// LS Electric XG5000 project: SEMICON_SORTER
// PLC DR32H

PROGRAM SIM_IO (task: 스캔 프로그램)

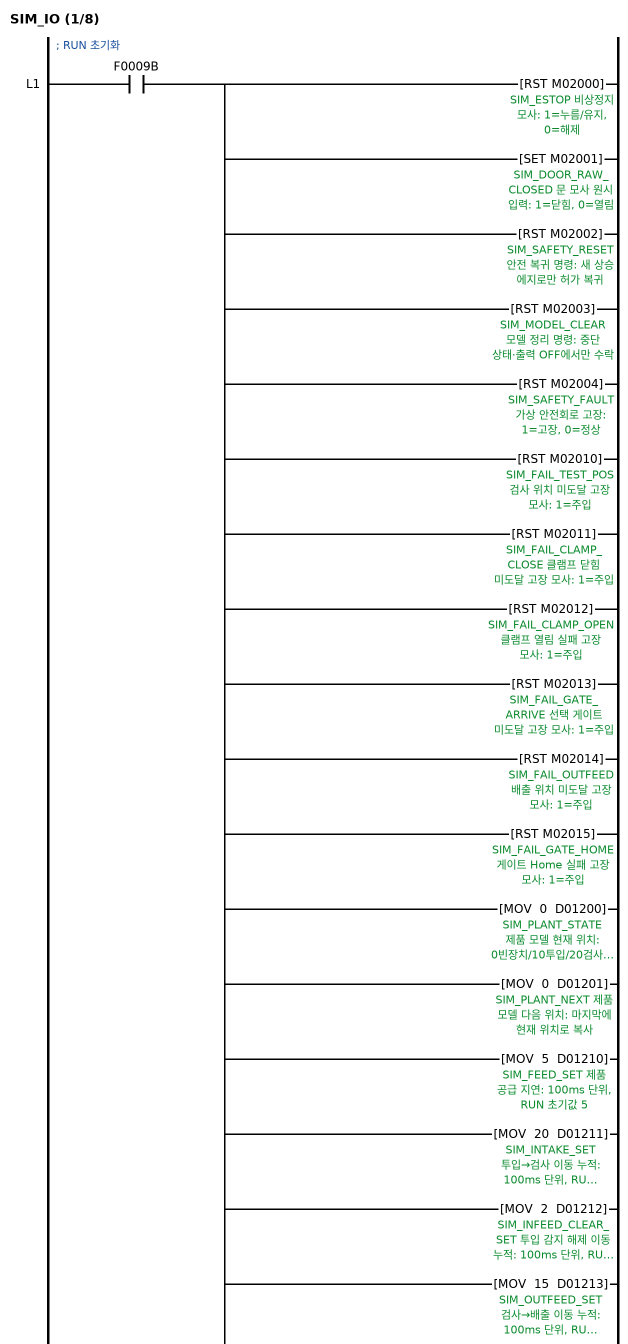

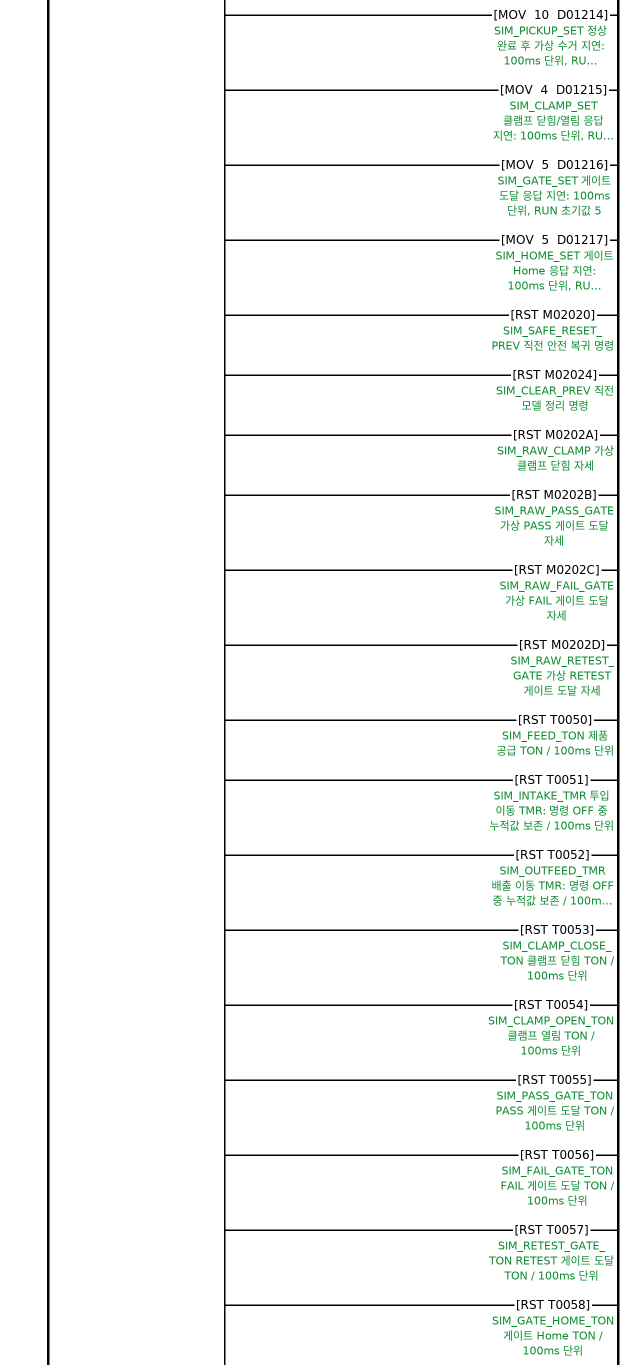

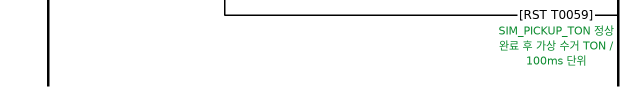
// RUN 초기화
; L1
LOAD      F0009B
RST       M02000	// SIM_ESTOP 비상정지 모사: 1=누름/유지, 0=해제
SET       M02001	// SIM_DOOR_RAW_CLOSED 문 모사 원시 입력: 1=닫힘, 0=열림
RST       M02002	// SIM_SAFETY_RESET 안전 복귀 명령: 새 상승 에지로만 허가 복귀
RST       M02003	// SIM_MODEL_CLEAR 모델 정리 명령: 중단 상태·출력 OFF에서만 수락
RST       M02004	// SIM_SAFETY_FAULT 가상 안전회로 고장: 1=고장, 0=정상
RST       M02010	// SIM_FAIL_TEST_POS 검사 위치 미도달 고장 모사: 1=주입
RST       M02011	// SIM_FAIL_CLAMP_CLOSE 클램프 닫힘 미도달 고장 모사: 1=주입
RST       M02012	// SIM_FAIL_CLAMP_OPEN 클램프 열림 실패 고장 모사: 1=주입
RST       M02013	// SIM_FAIL_GATE_ARRIVE 선택 게이트 미도달 고장 모사: 1=주입
RST       M02014	// SIM_FAIL_OUTFEED 배출 위치 미도달 고장 모사: 1=주입
RST       M02015	// SIM_FAIL_GATE_HOME 게이트 Home 실패 고장 모사: 1=주입
MOV       0 D01200	// SIM_PLANT_STATE 제품 모델 현재 위치: 0빈장치/10투입/20검사/30배출이송/40배출
MOV       0 D01201	// SIM_PLANT_NEXT 제품 모델 다음 위치: 마지막에 현재 위치로 복사
MOV       5 D01210	// SIM_FEED_SET 제품 공급 지연: 100ms 단위, RUN 초기값 5
MOV       20 D01211	// SIM_INTAKE_SET 투입→검사 이동 누적: 100ms 단위, RUN 초기값 20
MOV       2 D01212	// SIM_INFEED_CLEAR_SET 투입 감지 해제 이동 누적: 100ms 단위, RUN 초기값 2
MOV       15 D01213	// SIM_OUTFEED_SET 검사→배출 이동 누적: 100ms 단위, RUN 초기값 15
MOV       10 D01214	// SIM_PICKUP_SET 정상 완료 후 가상 수거 지연: 100ms 단위, RUN 초기값 10
MOV       4 D01215	// SIM_CLAMP_SET 클램프 닫힘/열림 응답 지연: 100ms 단위, RUN 초기값 4
MOV       5 D01216	// SIM_GATE_SET 게이트 도달 응답 지연: 100ms 단위, RUN 초기값 5
MOV       5 D01217	// SIM_HOME_SET 게이트 Home 응답 지연: 100ms 단위, RUN 초기값 5
RST       M02020	// SIM_SAFE_RESET_PREV 직전 안전 복귀 명령
RST       M02024	// SIM_CLEAR_PREV 직전 모델 정리 명령
RST       M0202A	// SIM_RAW_CLAMP 가상 클램프 닫힘 자세
RST       M0202B	// SIM_RAW_PASS_GATE 가상 PASS 게이트 도달 자세
RST       M0202C	// SIM_RAW_FAIL_GATE 가상 FAIL 게이트 도달 자세
RST       M0202D	// SIM_RAW_RETEST_GATE 가상 RETEST 게이트 도달 자세
RST       T0050	// SIM_FEED_TON 제품 공급 TON / 100ms 단위
RST       T0051	// SIM_INTAKE_TMR 투입 이동 TMR: 명령 OFF 중 누적값 보존 / 100ms 단위
RST       T0052	// SIM_OUTFEED_TMR 배출 이동 TMR: 명령 OFF 중 누적값 보존 / 100ms 단위
RST       T0053	// SIM_CLAMP_CLOSE_TON 클램프 닫힘 TON / 100ms 단위
RST       T0054	// SIM_CLAMP_OPEN_TON 클램프 열림 TON / 100ms 단위
RST       T0055	// SIM_PASS_GATE_TON PASS 게이트 도달 TON / 100ms 단위
RST       T0056	// SIM_FAIL_GATE_TON FAIL 게이트 도달 TON / 100ms 단위
RST       T0057	// SIM_RETEST_GATE_TON RETEST 게이트 도달 TON / 100ms 단위
RST       T0058	// SIM_GATE_HOME_TON 게이트 Home TON / 100ms 단위
RST       T0059	// SIM_PICKUP_TON 정상 완료 후 가상 수거 TON / 100ms 단위

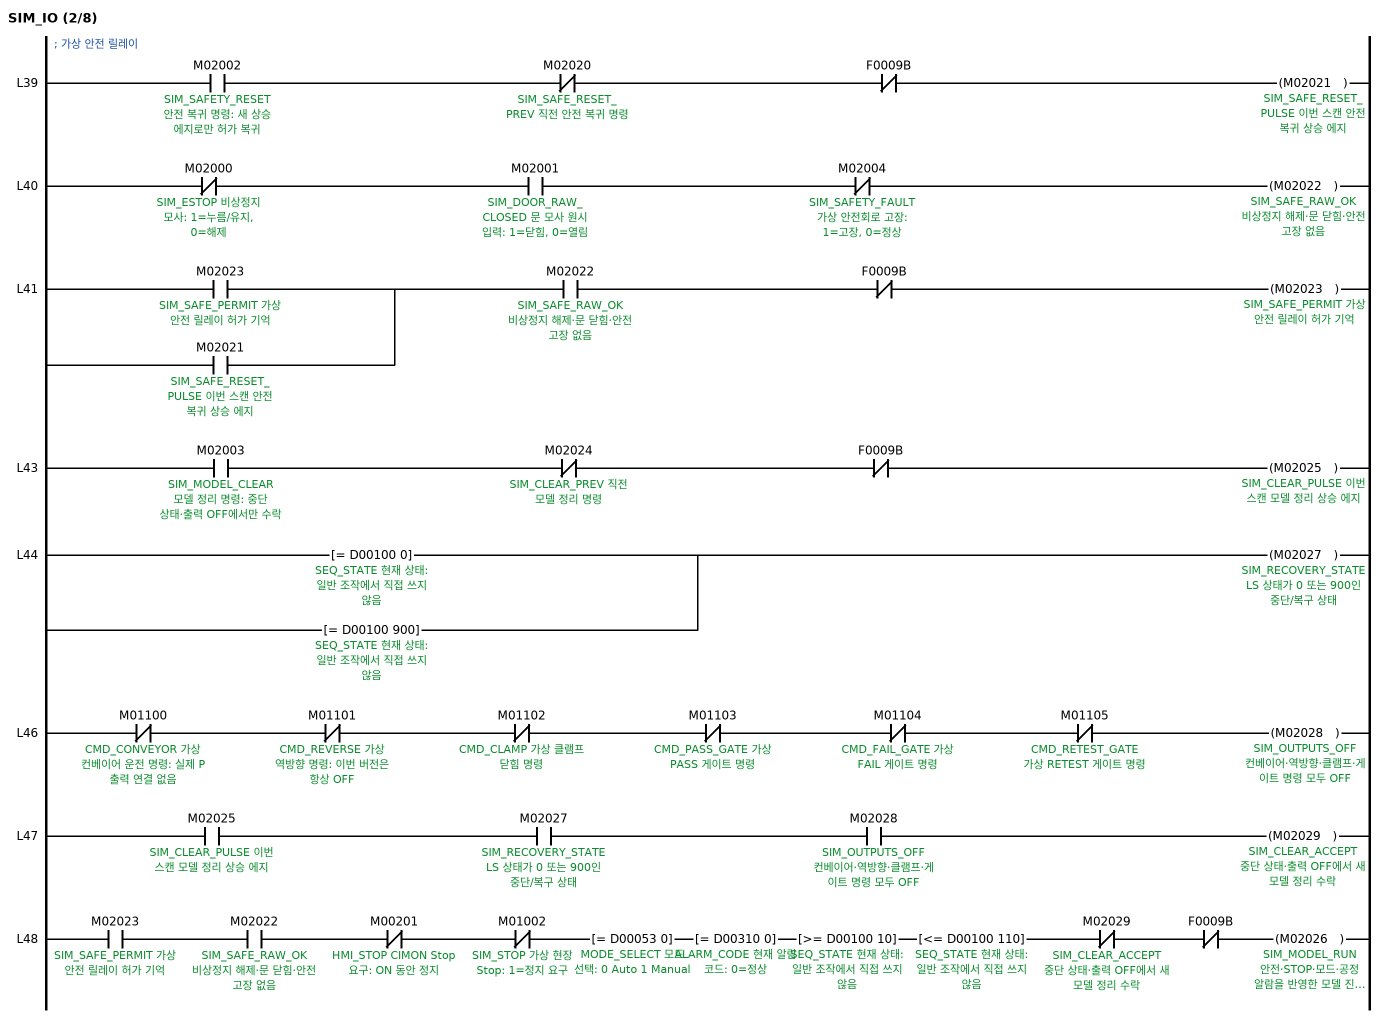
// 가상 안전 릴레이
; L39
LOAD      M02002	// SIM_SAFETY_RESET 안전 복귀 명령: 새 상승 에지로만 허가 복귀
AND NOT   M02020	// SIM_SAFE_RESET_PREV 직전 안전 복귀 명령
AND NOT   F0009B
OUT       M02021	// SIM_SAFE_RESET_PULSE 이번 스캔 안전 복귀 상승 에지
; L40
LOAD NOT  M02000	// SIM_ESTOP 비상정지 모사: 1=누름/유지, 0=해제
AND       M02001	// SIM_DOOR_RAW_CLOSED 문 모사 원시 입력: 1=닫힘, 0=열림
AND NOT   M02004	// SIM_SAFETY_FAULT 가상 안전회로 고장: 1=고장, 0=정상
OUT       M02022	// SIM_SAFE_RAW_OK 비상정지 해제·문 닫힘·안전 고장 없음
; L41
LOAD      M02023	// SIM_SAFE_PERMIT 가상 안전 릴레이 허가 기억
OR        M02021	// SIM_SAFE_RESET_PULSE 이번 스캔 안전 복귀 상승 에지
AND       M02022	// SIM_SAFE_RAW_OK 비상정지 해제·문 닫힘·안전 고장 없음
AND NOT   F0009B
OUT       M02023	// SIM_SAFE_PERMIT 가상 안전 릴레이 허가 기억
; L43
LOAD      M02003	// SIM_MODEL_CLEAR 모델 정리 명령: 중단 상태·출력 OFF에서만 수락
AND NOT   M02024	// SIM_CLEAR_PREV 직전 모델 정리 명령
AND NOT   F0009B
OUT       M02025	// SIM_CLEAR_PULSE 이번 스캔 모델 정리 상승 에지
; L44
LOAD=     D00100 0	// SEQ_STATE 현재 상태: 일반 조작에서 직접 쓰지 않음
OR=       D00100 900	// SEQ_STATE 현재 상태: 일반 조작에서 직접 쓰지 않음
OUT       M02027	// SIM_RECOVERY_STATE LS 상태가 0 또는 900인 중단/복구 상태
; L46
LOAD NOT  M01100	// CMD_CONVEYOR 가상 컨베이어 운전 명령: 실제 P 출력 연결 없음
AND NOT   M01101	// CMD_REVERSE 가상 역방향 명령: 이번 버전은 항상 OFF
AND NOT   M01102	// CMD_CLAMP 가상 클램프 닫힘 명령
AND NOT   M01103	// CMD_PASS_GATE 가상 PASS 게이트 명령
AND NOT   M01104	// CMD_FAIL_GATE 가상 FAIL 게이트 명령
AND NOT   M01105	// CMD_RETEST_GATE 가상 RETEST 게이트 명령
OUT       M02028	// SIM_OUTPUTS_OFF 컨베이어·역방향·클램프·게이트 명령 모두 OFF
; L47
LOAD      M02025	// SIM_CLEAR_PULSE 이번 스캔 모델 정리 상승 에지
AND       M02027	// SIM_RECOVERY_STATE LS 상태가 0 또는 900인 중단/복구 상태
AND       M02028	// SIM_OUTPUTS_OFF 컨베이어·역방향·클램프·게이트 명령 모두 OFF
OUT       M02029	// SIM_CLEAR_ACCEPT 중단 상태·출력 OFF에서 새 모델 정리 수락
; L48
LOAD      M02023	// SIM_SAFE_PERMIT 가상 안전 릴레이 허가 기억
AND       M02022	// SIM_SAFE_RAW_OK 비상정지 해제·문 닫힘·안전 고장 없음
AND NOT   M00201	// HMI_STOP CIMON Stop 요구: ON 동안 정지
AND NOT   M01002	// SIM_STOP 가상 현장 Stop: 1=정지 요구
AND=      D00053 0	// MODE_SELECT 모드 선택: 0 Auto 1 Manual
AND=      D00310 0	// ALARM_CODE 현재 알람 코드: 0=정상
AND>=     D00100 10	// SEQ_STATE 현재 상태: 일반 조작에서 직접 쓰지 않음
AND<=     D00100 110	// SEQ_STATE 현재 상태: 일반 조작에서 직접 쓰지 않음
AND NOT   M02029	// SIM_CLEAR_ACCEPT 중단 상태·출력 OFF에서 새 모델 정리 수락
AND NOT   F0009B
OUT       M02026	// SIM_MODEL_RUN 안전·STOP·모드·공정 알람을 반영한 모델 진행 허가

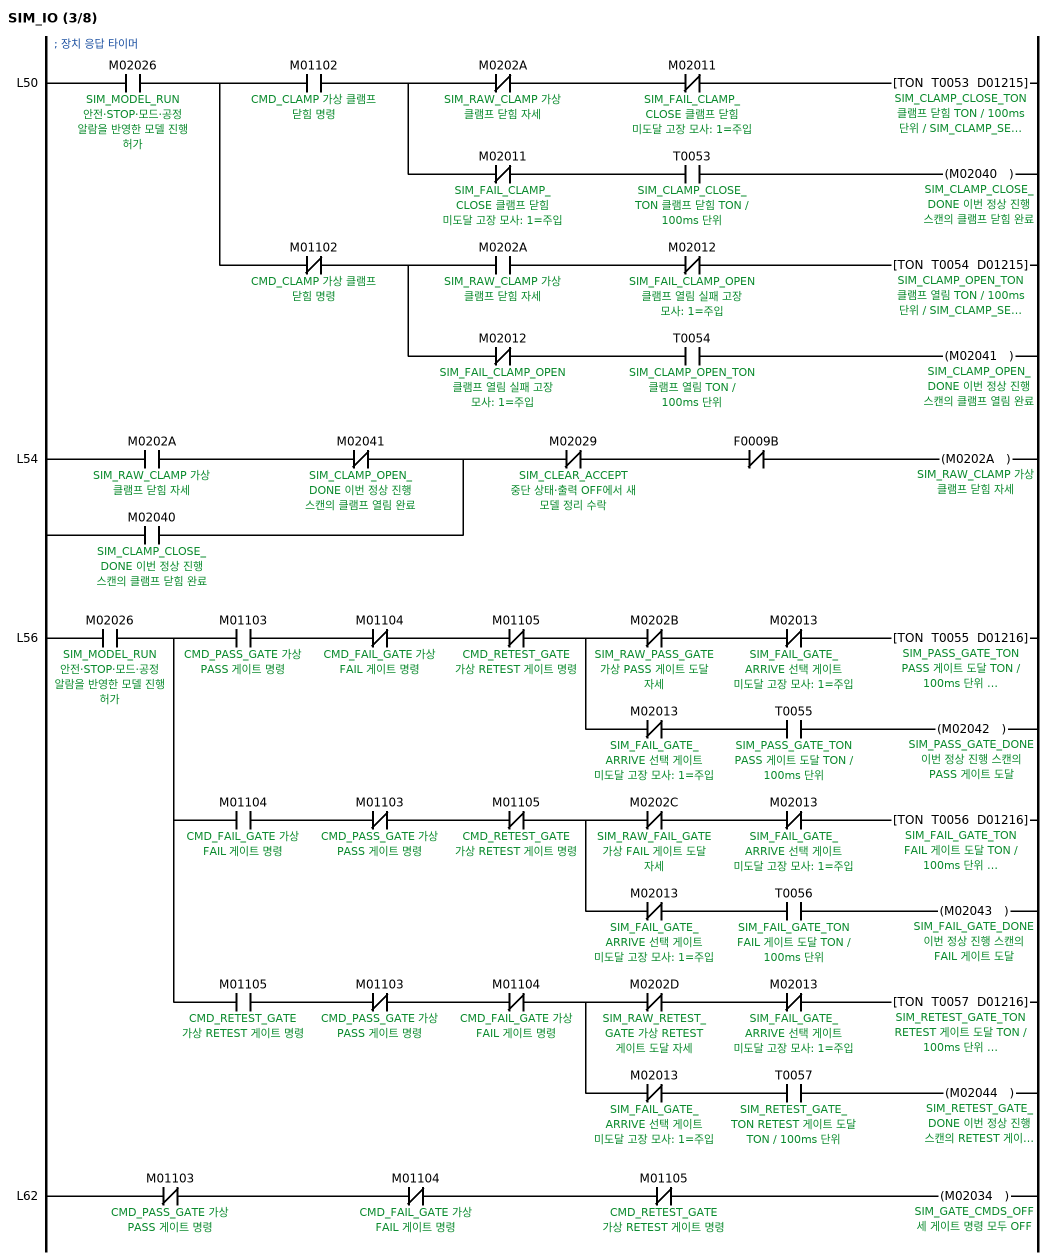
// 장치 응답 타이머
; L50
LOAD      M02026	// SIM_MODEL_RUN 안전·STOP·모드·공정 알람을 반영한 모델 진행 허가
MPUSH
AND       M01102	// CMD_CLAMP 가상 클램프 닫힘 명령
MPUSH
AND NOT   M0202A	// SIM_RAW_CLAMP 가상 클램프 닫힘 자세
AND NOT   M02011	// SIM_FAIL_CLAMP_CLOSE 클램프 닫힘 미도달 고장 모사: 1=주입
TON       T0053 D01215	// SIM_CLAMP_CLOSE_TON 클램프 닫힘 TON / 100ms 단위 / SIM_CLAMP_SET 클램프 닫힘/열림 응답 지연: 100ms 단위, RUN 초기값 4
MPOP
AND NOT   M02011	// SIM_FAIL_CLAMP_CLOSE 클램프 닫힘 미도달 고장 모사: 1=주입
AND       T0053	// SIM_CLAMP_CLOSE_TON 클램프 닫힘 TON / 100ms 단위
OUT       M02040	// SIM_CLAMP_CLOSE_DONE 이번 정상 진행 스캔의 클램프 닫힘 완료
MPOP
AND NOT   M01102	// CMD_CLAMP 가상 클램프 닫힘 명령
MPUSH
AND       M0202A	// SIM_RAW_CLAMP 가상 클램프 닫힘 자세
AND NOT   M02012	// SIM_FAIL_CLAMP_OPEN 클램프 열림 실패 고장 모사: 1=주입
TON       T0054 D01215	// SIM_CLAMP_OPEN_TON 클램프 열림 TON / 100ms 단위 / SIM_CLAMP_SET 클램프 닫힘/열림 응답 지연: 100ms 단위, RUN 초기값 4
MPOP
AND NOT   M02012	// SIM_FAIL_CLAMP_OPEN 클램프 열림 실패 고장 모사: 1=주입
AND       T0054	// SIM_CLAMP_OPEN_TON 클램프 열림 TON / 100ms 단위
OUT       M02041	// SIM_CLAMP_OPEN_DONE 이번 정상 진행 스캔의 클램프 열림 완료
; L54
LOAD      M0202A	// SIM_RAW_CLAMP 가상 클램프 닫힘 자세
AND NOT   M02041	// SIM_CLAMP_OPEN_DONE 이번 정상 진행 스캔의 클램프 열림 완료
OR        M02040	// SIM_CLAMP_CLOSE_DONE 이번 정상 진행 스캔의 클램프 닫힘 완료
AND NOT   M02029	// SIM_CLEAR_ACCEPT 중단 상태·출력 OFF에서 새 모델 정리 수락
AND NOT   F0009B
OUT       M0202A	// SIM_RAW_CLAMP 가상 클램프 닫힘 자세
; L56
LOAD      M02026	// SIM_MODEL_RUN 안전·STOP·모드·공정 알람을 반영한 모델 진행 허가
MPUSH
AND       M01103	// CMD_PASS_GATE 가상 PASS 게이트 명령
AND NOT   M01104	// CMD_FAIL_GATE 가상 FAIL 게이트 명령
AND NOT   M01105	// CMD_RETEST_GATE 가상 RETEST 게이트 명령
MPUSH
AND NOT   M0202B	// SIM_RAW_PASS_GATE 가상 PASS 게이트 도달 자세
AND NOT   M02013	// SIM_FAIL_GATE_ARRIVE 선택 게이트 미도달 고장 모사: 1=주입
TON       T0055 D01216	// SIM_PASS_GATE_TON PASS 게이트 도달 TON / 100ms 단위 / SIM_GATE_SET 게이트 도달 응답 지연: 100ms 단위, RUN 초기값 5
MPOP
AND NOT   M02013	// SIM_FAIL_GATE_ARRIVE 선택 게이트 미도달 고장 모사: 1=주입
AND       T0055	// SIM_PASS_GATE_TON PASS 게이트 도달 TON / 100ms 단위
OUT       M02042	// SIM_PASS_GATE_DONE 이번 정상 진행 스캔의 PASS 게이트 도달
MLOAD
AND       M01104	// CMD_FAIL_GATE 가상 FAIL 게이트 명령
AND NOT   M01103	// CMD_PASS_GATE 가상 PASS 게이트 명령
AND NOT   M01105	// CMD_RETEST_GATE 가상 RETEST 게이트 명령
MPUSH
AND NOT   M0202C	// SIM_RAW_FAIL_GATE 가상 FAIL 게이트 도달 자세
AND NOT   M02013	// SIM_FAIL_GATE_ARRIVE 선택 게이트 미도달 고장 모사: 1=주입
TON       T0056 D01216	// SIM_FAIL_GATE_TON FAIL 게이트 도달 TON / 100ms 단위 / SIM_GATE_SET 게이트 도달 응답 지연: 100ms 단위, RUN 초기값 5
MPOP
AND NOT   M02013	// SIM_FAIL_GATE_ARRIVE 선택 게이트 미도달 고장 모사: 1=주입
AND       T0056	// SIM_FAIL_GATE_TON FAIL 게이트 도달 TON / 100ms 단위
OUT       M02043	// SIM_FAIL_GATE_DONE 이번 정상 진행 스캔의 FAIL 게이트 도달
MPOP
AND       M01105	// CMD_RETEST_GATE 가상 RETEST 게이트 명령
AND NOT   M01103	// CMD_PASS_GATE 가상 PASS 게이트 명령
AND NOT   M01104	// CMD_FAIL_GATE 가상 FAIL 게이트 명령
MPUSH
AND NOT   M0202D	// SIM_RAW_RETEST_GATE 가상 RETEST 게이트 도달 자세
AND NOT   M02013	// SIM_FAIL_GATE_ARRIVE 선택 게이트 미도달 고장 모사: 1=주입
TON       T0057 D01216	// SIM_RETEST_GATE_TON RETEST 게이트 도달 TON / 100ms 단위 / SIM_GATE_SET 게이트 도달 응답 지연: 100ms 단위, RUN 초기값 5
MPOP
AND NOT   M02013	// SIM_FAIL_GATE_ARRIVE 선택 게이트 미도달 고장 모사: 1=주입
AND       T0057	// SIM_RETEST_GATE_TON RETEST 게이트 도달 TON / 100ms 단위
OUT       M02044	// SIM_RETEST_GATE_DONE 이번 정상 진행 스캔의 RETEST 게이트 도달
; L62
LOAD NOT  M01103	// CMD_PASS_GATE 가상 PASS 게이트 명령
AND NOT   M01104	// CMD_FAIL_GATE 가상 FAIL 게이트 명령
AND NOT   M01105	// CMD_RETEST_GATE 가상 RETEST 게이트 명령
OUT       M02034	// SIM_GATE_CMDS_OFF 세 게이트 명령 모두 OFF

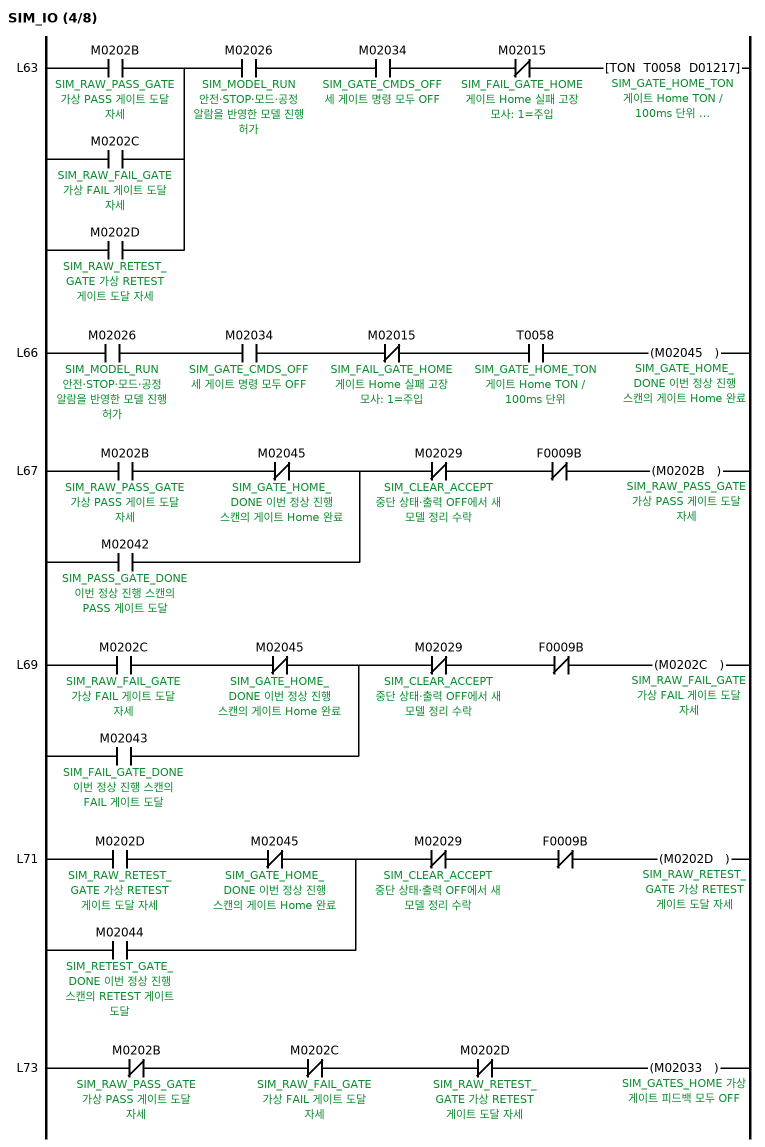
; L63
LOAD      M0202B	// SIM_RAW_PASS_GATE 가상 PASS 게이트 도달 자세
OR        M0202C	// SIM_RAW_FAIL_GATE 가상 FAIL 게이트 도달 자세
OR        M0202D	// SIM_RAW_RETEST_GATE 가상 RETEST 게이트 도달 자세
AND       M02026	// SIM_MODEL_RUN 안전·STOP·모드·공정 알람을 반영한 모델 진행 허가
AND       M02034	// SIM_GATE_CMDS_OFF 세 게이트 명령 모두 OFF
AND NOT   M02015	// SIM_FAIL_GATE_HOME 게이트 Home 실패 고장 모사: 1=주입
TON       T0058 D01217	// SIM_GATE_HOME_TON 게이트 Home TON / 100ms 단위 / SIM_HOME_SET 게이트 Home 응답 지연: 100ms 단위, RUN 초기값 5
; L66
LOAD      M02026	// SIM_MODEL_RUN 안전·STOP·모드·공정 알람을 반영한 모델 진행 허가
AND       M02034	// SIM_GATE_CMDS_OFF 세 게이트 명령 모두 OFF
AND NOT   M02015	// SIM_FAIL_GATE_HOME 게이트 Home 실패 고장 모사: 1=주입
AND       T0058	// SIM_GATE_HOME_TON 게이트 Home TON / 100ms 단위
OUT       M02045	// SIM_GATE_HOME_DONE 이번 정상 진행 스캔의 게이트 Home 완료
; L67
LOAD      M0202B	// SIM_RAW_PASS_GATE 가상 PASS 게이트 도달 자세
AND NOT   M02045	// SIM_GATE_HOME_DONE 이번 정상 진행 스캔의 게이트 Home 완료
OR        M02042	// SIM_PASS_GATE_DONE 이번 정상 진행 스캔의 PASS 게이트 도달
AND NOT   M02029	// SIM_CLEAR_ACCEPT 중단 상태·출력 OFF에서 새 모델 정리 수락
AND NOT   F0009B
OUT       M0202B	// SIM_RAW_PASS_GATE 가상 PASS 게이트 도달 자세
; L69
LOAD      M0202C	// SIM_RAW_FAIL_GATE 가상 FAIL 게이트 도달 자세
AND NOT   M02045	// SIM_GATE_HOME_DONE 이번 정상 진행 스캔의 게이트 Home 완료
OR        M02043	// SIM_FAIL_GATE_DONE 이번 정상 진행 스캔의 FAIL 게이트 도달
AND NOT   M02029	// SIM_CLEAR_ACCEPT 중단 상태·출력 OFF에서 새 모델 정리 수락
AND NOT   F0009B
OUT       M0202C	// SIM_RAW_FAIL_GATE 가상 FAIL 게이트 도달 자세
; L71
LOAD      M0202D	// SIM_RAW_RETEST_GATE 가상 RETEST 게이트 도달 자세
AND NOT   M02045	// SIM_GATE_HOME_DONE 이번 정상 진행 스캔의 게이트 Home 완료
OR        M02044	// SIM_RETEST_GATE_DONE 이번 정상 진행 스캔의 RETEST 게이트 도달
AND NOT   M02029	// SIM_CLEAR_ACCEPT 중단 상태·출력 OFF에서 새 모델 정리 수락
AND NOT   F0009B
OUT       M0202D	// SIM_RAW_RETEST_GATE 가상 RETEST 게이트 도달 자세
; L73
LOAD NOT  M0202B	// SIM_RAW_PASS_GATE 가상 PASS 게이트 도달 자세
AND NOT   M0202C	// SIM_RAW_FAIL_GATE 가상 FAIL 게이트 도달 자세
AND NOT   M0202D	// SIM_RAW_RETEST_GATE 가상 RETEST 게이트 도달 자세
OUT       M02033	// SIM_GATES_HOME 가상 게이트 피드백 모두 OFF

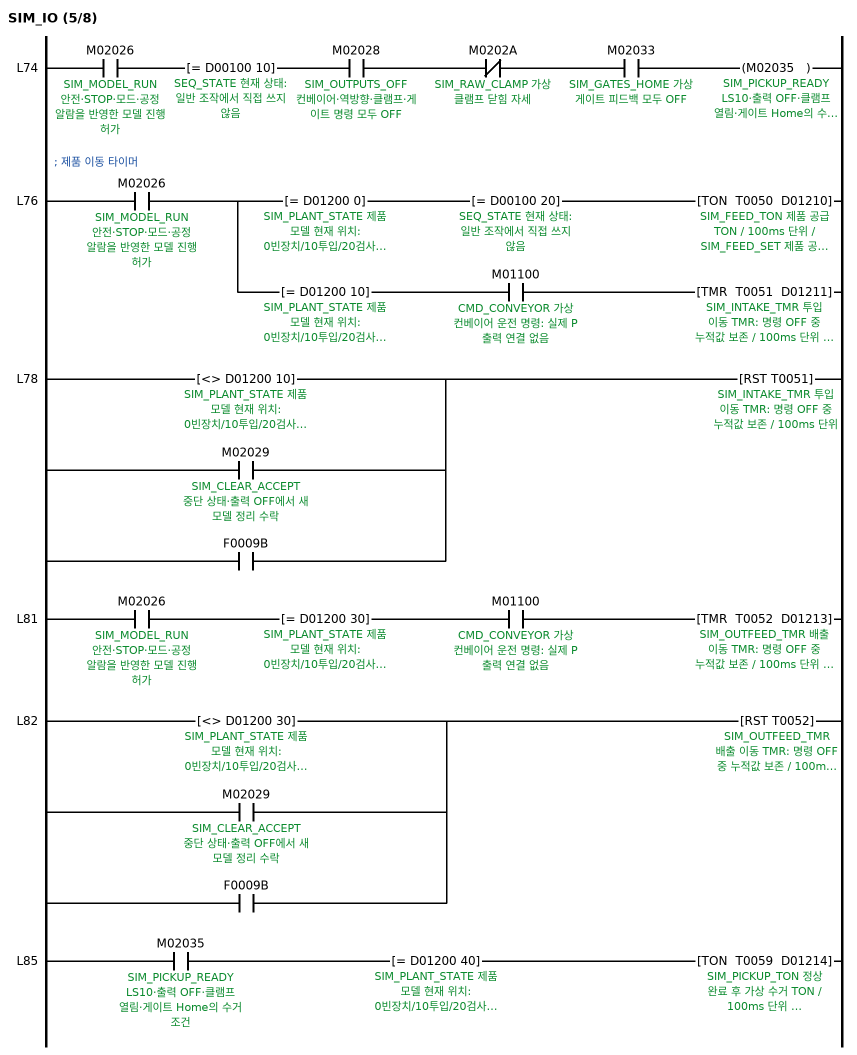
; L74
LOAD      M02026	// SIM_MODEL_RUN 안전·STOP·모드·공정 알람을 반영한 모델 진행 허가
AND=      D00100 10	// SEQ_STATE 현재 상태: 일반 조작에서 직접 쓰지 않음
AND       M02028	// SIM_OUTPUTS_OFF 컨베이어·역방향·클램프·게이트 명령 모두 OFF
AND NOT   M0202A	// SIM_RAW_CLAMP 가상 클램프 닫힘 자세
AND       M02033	// SIM_GATES_HOME 가상 게이트 피드백 모두 OFF
OUT       M02035	// SIM_PICKUP_READY LS10·출력 OFF·클램프 열림·게이트 Home의 수거 조건
// 제품 이동 타이머
; L76
LOAD      M02026	// SIM_MODEL_RUN 안전·STOP·모드·공정 알람을 반영한 모델 진행 허가
MPUSH
AND=      D01200 0	// SIM_PLANT_STATE 제품 모델 현재 위치: 0빈장치/10투입/20검사/30배출이송/40배출
AND=      D00100 20	// SEQ_STATE 현재 상태: 일반 조작에서 직접 쓰지 않음
TON       T0050 D01210	// SIM_FEED_TON 제품 공급 TON / 100ms 단위 / SIM_FEED_SET 제품 공급 지연: 100ms 단위, RUN 초기값 5
MPOP
AND=      D01200 10	// SIM_PLANT_STATE 제품 모델 현재 위치: 0빈장치/10투입/20검사/30배출이송/40배출
AND       M01100	// CMD_CONVEYOR 가상 컨베이어 운전 명령: 실제 P 출력 연결 없음
TMR       T0051 D01211	// SIM_INTAKE_TMR 투입 이동 TMR: 명령 OFF 중 누적값 보존 / 100ms 단위 / SIM_INTAKE_SET 투입→검사 이동 누적: 100ms 단위, RUN 초기값 20
; L78
LOAD<>    D01200 10	// SIM_PLANT_STATE 제품 모델 현재 위치: 0빈장치/10투입/20검사/30배출이송/40배출
OR        M02029	// SIM_CLEAR_ACCEPT 중단 상태·출력 OFF에서 새 모델 정리 수락
OR        F0009B
RST       T0051	// SIM_INTAKE_TMR 투입 이동 TMR: 명령 OFF 중 누적값 보존 / 100ms 단위
; L81
LOAD      M02026	// SIM_MODEL_RUN 안전·STOP·모드·공정 알람을 반영한 모델 진행 허가
AND=      D01200 30	// SIM_PLANT_STATE 제품 모델 현재 위치: 0빈장치/10투입/20검사/30배출이송/40배출
AND       M01100	// CMD_CONVEYOR 가상 컨베이어 운전 명령: 실제 P 출력 연결 없음
TMR       T0052 D01213	// SIM_OUTFEED_TMR 배출 이동 TMR: 명령 OFF 중 누적값 보존 / 100ms 단위 / SIM_OUTFEED_SET 검사→배출 이동 누적: 100ms 단위, RUN 초기값 15
; L82
LOAD<>    D01200 30	// SIM_PLANT_STATE 제품 모델 현재 위치: 0빈장치/10투입/20검사/30배출이송/40배출
OR        M02029	// SIM_CLEAR_ACCEPT 중단 상태·출력 OFF에서 새 모델 정리 수락
OR        F0009B
RST       T0052	// SIM_OUTFEED_TMR 배출 이동 TMR: 명령 OFF 중 누적값 보존 / 100ms 단위
; L85
LOAD      M02035	// SIM_PICKUP_READY LS10·출력 OFF·클램프 열림·게이트 Home의 수거 조건
AND=      D01200 40	// SIM_PLANT_STATE 제품 모델 현재 위치: 0빈장치/10투입/20검사/30배출이송/40배출
TON       T0059 D01214	// SIM_PICKUP_TON 정상 완료 후 가상 수거 TON / 100ms 단위 / SIM_PICKUP_SET 정상 완료 후 가상 수거 지연: 100ms 단위, RUN 초기값 10

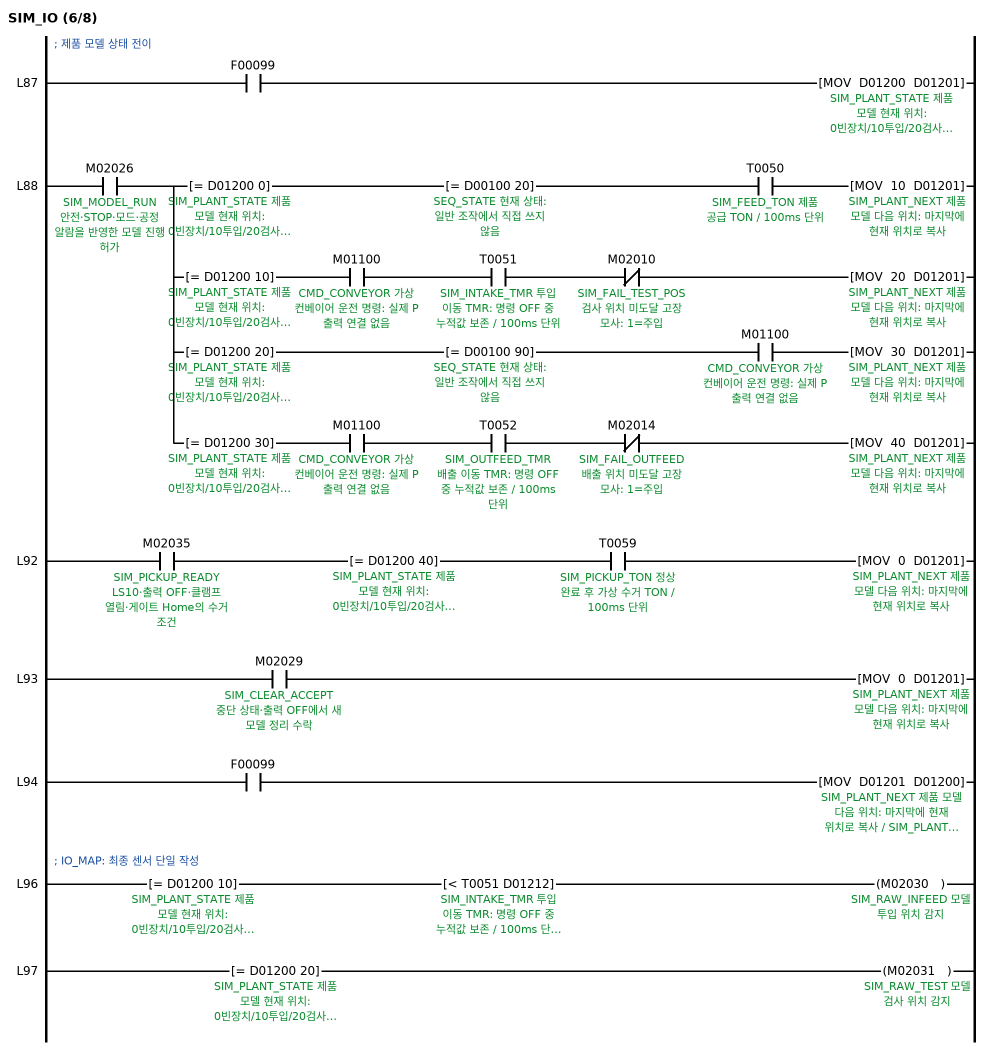
// 제품 모델 상태 전이
; L87
LOAD      F00099
MOV       D01200 D01201	// SIM_PLANT_STATE 제품 모델 현재 위치: 0빈장치/10투입/20검사/30배출이송/40배출 / SIM_PLANT_NEXT 제품 모델 다음 위치: 마지막에 현재 위치로 복사
; L88
LOAD      M02026	// SIM_MODEL_RUN 안전·STOP·모드·공정 알람을 반영한 모델 진행 허가
MPUSH
AND=      D01200 0	// SIM_PLANT_STATE 제품 모델 현재 위치: 0빈장치/10투입/20검사/30배출이송/40배출
AND=      D00100 20	// SEQ_STATE 현재 상태: 일반 조작에서 직접 쓰지 않음
AND       T0050	// SIM_FEED_TON 제품 공급 TON / 100ms 단위
MOV       10 D01201	// SIM_PLANT_NEXT 제품 모델 다음 위치: 마지막에 현재 위치로 복사
MLOAD
AND=      D01200 10	// SIM_PLANT_STATE 제품 모델 현재 위치: 0빈장치/10투입/20검사/30배출이송/40배출
AND       M01100	// CMD_CONVEYOR 가상 컨베이어 운전 명령: 실제 P 출력 연결 없음
AND       T0051	// SIM_INTAKE_TMR 투입 이동 TMR: 명령 OFF 중 누적값 보존 / 100ms 단위
AND NOT   M02010	// SIM_FAIL_TEST_POS 검사 위치 미도달 고장 모사: 1=주입
MOV       20 D01201	// SIM_PLANT_NEXT 제품 모델 다음 위치: 마지막에 현재 위치로 복사
MLOAD
AND=      D01200 20	// SIM_PLANT_STATE 제품 모델 현재 위치: 0빈장치/10투입/20검사/30배출이송/40배출
AND=      D00100 90	// SEQ_STATE 현재 상태: 일반 조작에서 직접 쓰지 않음
AND       M01100	// CMD_CONVEYOR 가상 컨베이어 운전 명령: 실제 P 출력 연결 없음
MOV       30 D01201	// SIM_PLANT_NEXT 제품 모델 다음 위치: 마지막에 현재 위치로 복사
MPOP
AND=      D01200 30	// SIM_PLANT_STATE 제품 모델 현재 위치: 0빈장치/10투입/20검사/30배출이송/40배출
AND       M01100	// CMD_CONVEYOR 가상 컨베이어 운전 명령: 실제 P 출력 연결 없음
AND       T0052	// SIM_OUTFEED_TMR 배출 이동 TMR: 명령 OFF 중 누적값 보존 / 100ms 단위
AND NOT   M02014	// SIM_FAIL_OUTFEED 배출 위치 미도달 고장 모사: 1=주입
MOV       40 D01201	// SIM_PLANT_NEXT 제품 모델 다음 위치: 마지막에 현재 위치로 복사
; L92
LOAD      M02035	// SIM_PICKUP_READY LS10·출력 OFF·클램프 열림·게이트 Home의 수거 조건
AND=      D01200 40	// SIM_PLANT_STATE 제품 모델 현재 위치: 0빈장치/10투입/20검사/30배출이송/40배출
AND       T0059	// SIM_PICKUP_TON 정상 완료 후 가상 수거 TON / 100ms 단위
MOV       0 D01201	// SIM_PLANT_NEXT 제품 모델 다음 위치: 마지막에 현재 위치로 복사
; L93
LOAD      M02029	// SIM_CLEAR_ACCEPT 중단 상태·출력 OFF에서 새 모델 정리 수락
MOV       0 D01201	// SIM_PLANT_NEXT 제품 모델 다음 위치: 마지막에 현재 위치로 복사
; L94
LOAD      F00099
MOV       D01201 D01200	// SIM_PLANT_NEXT 제품 모델 다음 위치: 마지막에 현재 위치로 복사 / SIM_PLANT_STATE 제품 모델 현재 위치: 0빈장치/10투입/20검사/30배출이송/40배출
// IO_MAP: 최종 센서 단일 작성
; L96
LOAD=     D01200 10	// SIM_PLANT_STATE 제품 모델 현재 위치: 0빈장치/10투입/20검사/30배출이송/40배출
AND<      T0051 D01212	// SIM_INTAKE_TMR 투입 이동 TMR: 명령 OFF 중 누적값 보존 / 100ms 단위 / SIM_INFEED_CLEAR_SET 투입 감지 해제 이동 누적: 100ms 단위, RUN 초기값 2
OUT       M02030	// SIM_RAW_INFEED 모델 투입 위치 감지
; L97
LOAD=     D01200 20	// SIM_PLANT_STATE 제품 모델 현재 위치: 0빈장치/10투입/20검사/30배출이송/40배출
OUT       M02031	// SIM_RAW_TEST 모델 검사 위치 감지

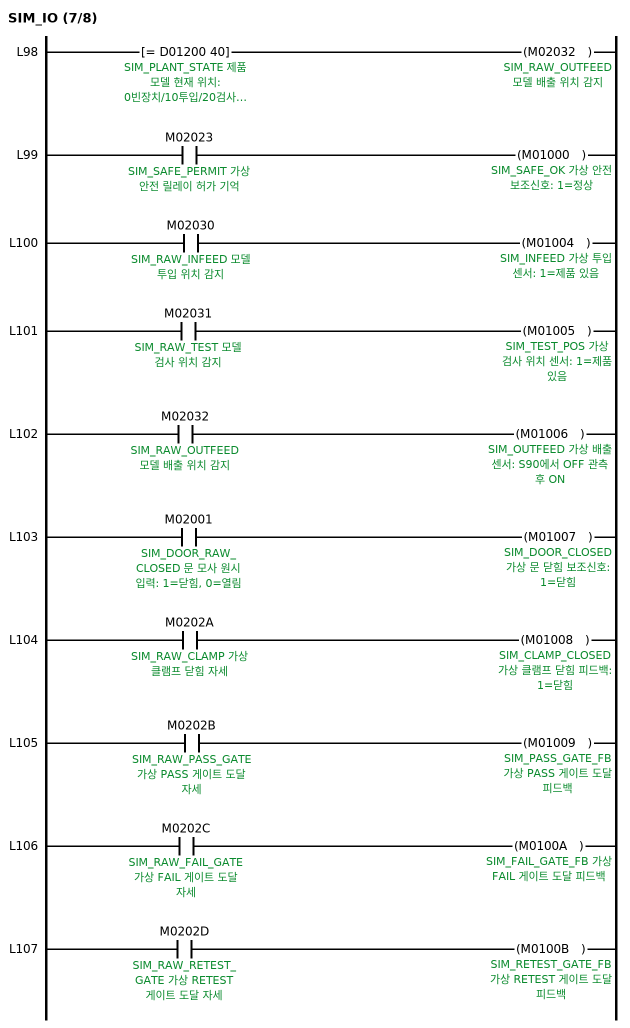
; L98
LOAD=     D01200 40	// SIM_PLANT_STATE 제품 모델 현재 위치: 0빈장치/10투입/20검사/30배출이송/40배출
OUT       M02032	// SIM_RAW_OUTFEED 모델 배출 위치 감지
; L99
LOAD      M02023	// SIM_SAFE_PERMIT 가상 안전 릴레이 허가 기억
OUT       M01000	// SIM_SAFE_OK 가상 안전 보조신호: 1=정상
; L100
LOAD      M02030	// SIM_RAW_INFEED 모델 투입 위치 감지
OUT       M01004	// SIM_INFEED 가상 투입 센서: 1=제품 있음
; L101
LOAD      M02031	// SIM_RAW_TEST 모델 검사 위치 감지
OUT       M01005	// SIM_TEST_POS 가상 검사 위치 센서: 1=제품 있음
; L102
LOAD      M02032	// SIM_RAW_OUTFEED 모델 배출 위치 감지
OUT       M01006	// SIM_OUTFEED 가상 배출 센서: S90에서 OFF 관측 후 ON
; L103
LOAD      M02001	// SIM_DOOR_RAW_CLOSED 문 모사 원시 입력: 1=닫힘, 0=열림
OUT       M01007	// SIM_DOOR_CLOSED 가상 문 닫힘 보조신호: 1=닫힘
; L104
LOAD      M0202A	// SIM_RAW_CLAMP 가상 클램프 닫힘 자세
OUT       M01008	// SIM_CLAMP_CLOSED 가상 클램프 닫힘 피드백: 1=닫힘
; L105
LOAD      M0202B	// SIM_RAW_PASS_GATE 가상 PASS 게이트 도달 자세
OUT       M01009	// SIM_PASS_GATE_FB 가상 PASS 게이트 도달 피드백
; L106
LOAD      M0202C	// SIM_RAW_FAIL_GATE 가상 FAIL 게이트 도달 자세
OUT       M0100A	// SIM_FAIL_GATE_FB 가상 FAIL 게이트 도달 피드백
; L107
LOAD      M0202D	// SIM_RAW_RETEST_GATE 가상 RETEST 게이트 도달 자세
OUT       M0100B	// SIM_RETEST_GATE_FB 가상 RETEST 게이트 도달 피드백

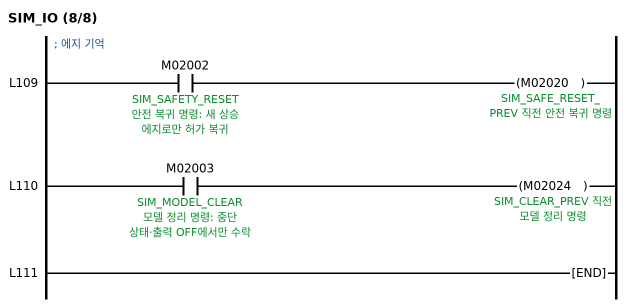
// 에지 기억
; L109
LOAD      M02002	// SIM_SAFETY_RESET 안전 복귀 명령: 새 상승 에지로만 허가 복귀
OUT       M02020	// SIM_SAFE_RESET_PREV 직전 안전 복귀 명령
; L110
LOAD      M02003	// SIM_MODEL_CLEAR 모델 정리 명령: 중단 상태·출력 OFF에서만 수락
OUT       M02024	// SIM_CLEAR_PREV 직전 모델 정리 명령
; L111
END

PROGRAM MAIN (task: 스캔 프로그램)

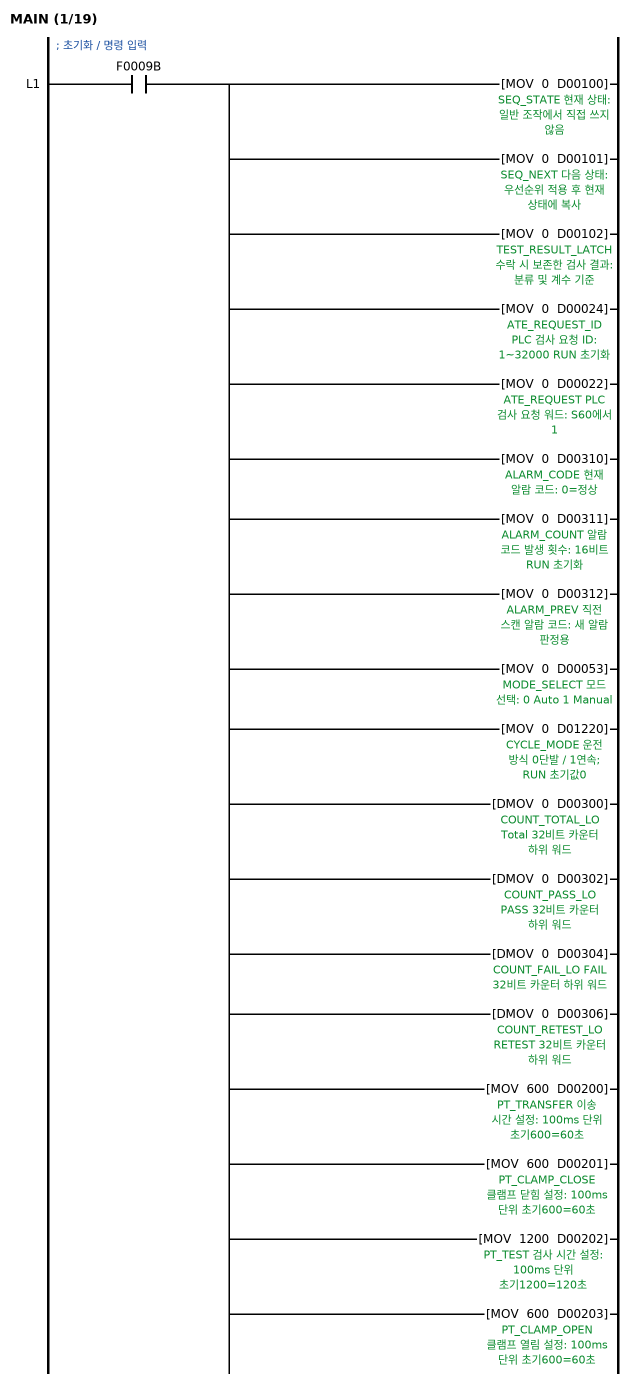

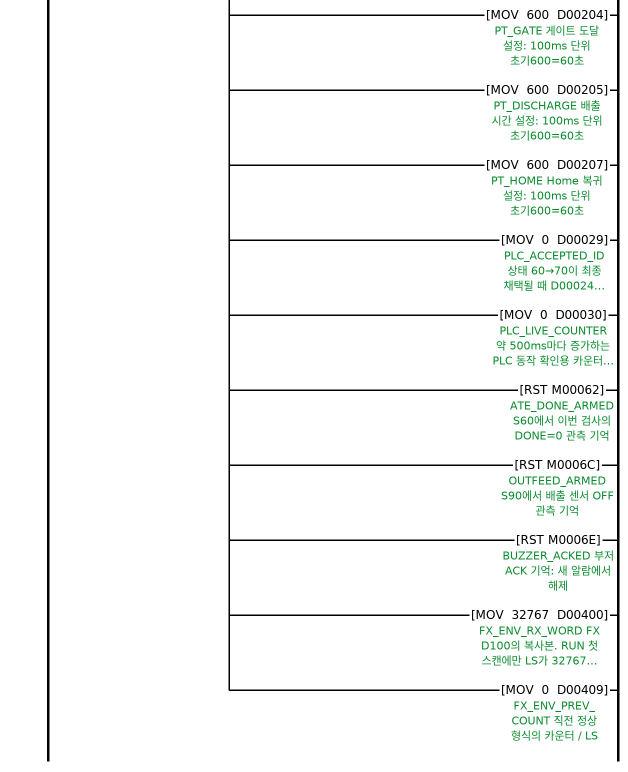
// 초기화 / 명령 입력
; L1
LOAD      F0009B
MOV       0 D00100	// SEQ_STATE 현재 상태: 일반 조작에서 직접 쓰지 않음
MOV       0 D00101	// SEQ_NEXT 다음 상태: 우선순위 적용 후 현재 상태에 복사
MOV       0 D00102	// TEST_RESULT_LATCH 수락 시 보존한 검사 결과: 분류 및 계수 기준
MOV       0 D00024	// ATE_REQUEST_ID PLC 검사 요청 ID: 1~32000 RUN 초기화
MOV       0 D00022	// ATE_REQUEST PLC 검사 요청 워드: S60에서 1
MOV       0 D00310	// ALARM_CODE 현재 알람 코드: 0=정상
MOV       0 D00311	// ALARM_COUNT 알람 코드 발생 횟수: 16비트 RUN 초기화
MOV       0 D00312	// ALARM_PREV 직전 스캔 알람 코드: 새 알람 판정용
MOV       0 D00053	// MODE_SELECT 모드 선택: 0 Auto 1 Manual
MOV       0 D01220	// CYCLE_MODE 운전 방식 0단발 / 1연속; RUN 초기값0
DMOV      0 D00300	// COUNT_TOTAL_LO Total 32비트 카운터 하위 워드
DMOV      0 D00302	// COUNT_PASS_LO PASS 32비트 카운터 하위 워드
DMOV      0 D00304	// COUNT_FAIL_LO FAIL 32비트 카운터 하위 워드
DMOV      0 D00306	// COUNT_RETEST_LO RETEST 32비트 카운터 하위 워드
MOV       600 D00200	// PT_TRANSFER 이송 시간 설정: 100ms 단위 초기600=60초
MOV       600 D00201	// PT_CLAMP_CLOSE 클램프 닫힘 설정: 100ms 단위 초기600=60초
MOV       1200 D00202	// PT_TEST 검사 시간 설정: 100ms 단위 초기1200=120초
MOV       600 D00203	// PT_CLAMP_OPEN 클램프 열림 설정: 100ms 단위 초기600=60초
MOV       600 D00204	// PT_GATE 게이트 도달 설정: 100ms 단위 초기600=60초
MOV       600 D00205	// PT_DISCHARGE 배출 시간 설정: 100ms 단위 초기600=60초
MOV       600 D00207	// PT_HOME Home 복귀 설정: 100ms 단위 초기600=60초
MOV       0 D00029	// PLC_ACCEPTED_ID 상태 60→70이 최종 채택될 때 D00024를 보존한 번호
MOV       0 D00030	// PLC_LIVE_COUNTER 약 500ms마다 증가하는 PLC 동작 확인용 카운터, 0~32000
RST       M00062	// ATE_DONE_ARMED S60에서 이번 검사의 DONE=0 관측 기억
RST       M0006C	// OUTFEED_ARMED S90에서 배출 센서 OFF 관측 기억
RST       M0006E	// BUZZER_ACKED 부저 ACK 기억: 새 알람에서 해제
MOV       32767 D00400	// FX_ENV_RX_WORD FX D100의 복사본. RUN 첫 스캔에만 LS가 32767로 초기화. 이후 모의시험 작업자 또는 CIMON 한 곳이 기록
MOV       0 D00409	// FX_ENV_PREV_COUNT 직전 정상 형식의 카운터 / LS

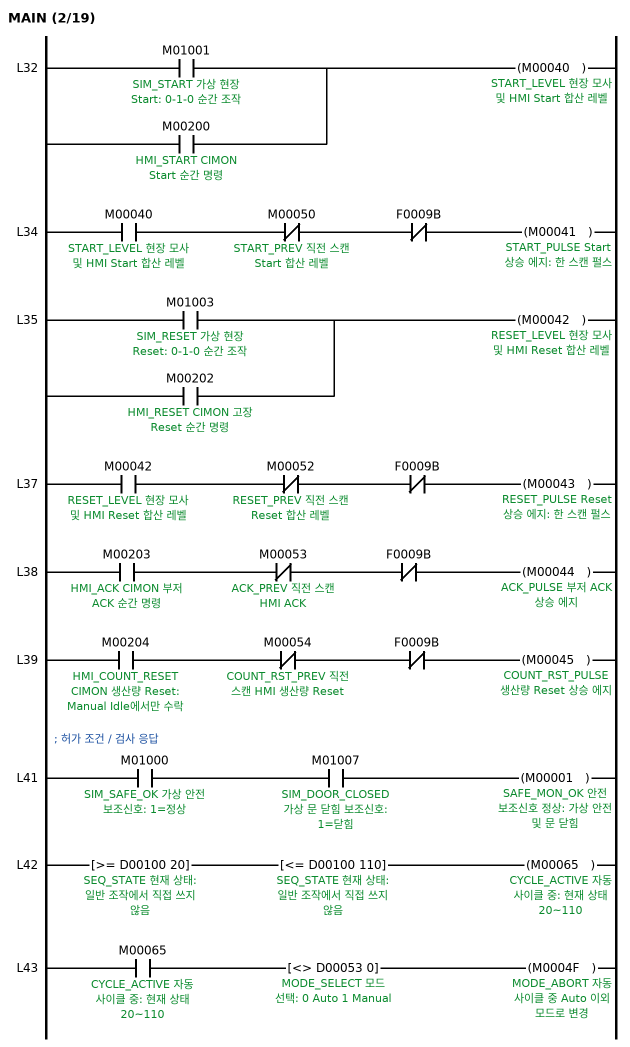
; L32
LOAD      M01001	// SIM_START 가상 현장 Start: 0-1-0 순간 조작
OR        M00200	// HMI_START CIMON Start 순간 명령
OUT       M00040	// START_LEVEL 현장 모사 및 HMI Start 합산 레벨
; L34
LOAD      M00040	// START_LEVEL 현장 모사 및 HMI Start 합산 레벨
AND NOT   M00050	// START_PREV 직전 스캔 Start 합산 레벨
AND NOT   F0009B
OUT       M00041	// START_PULSE Start 상승 에지: 한 스캔 펄스
; L35
LOAD      M01003	// SIM_RESET 가상 현장 Reset: 0-1-0 순간 조작
OR        M00202	// HMI_RESET CIMON 고장 Reset 순간 명령
OUT       M00042	// RESET_LEVEL 현장 모사 및 HMI Reset 합산 레벨
; L37
LOAD      M00042	// RESET_LEVEL 현장 모사 및 HMI Reset 합산 레벨
AND NOT   M00052	// RESET_PREV 직전 스캔 Reset 합산 레벨
AND NOT   F0009B
OUT       M00043	// RESET_PULSE Reset 상승 에지: 한 스캔 펄스
; L38
LOAD      M00203	// HMI_ACK CIMON 부저 ACK 순간 명령
AND NOT   M00053	// ACK_PREV 직전 스캔 HMI ACK
AND NOT   F0009B
OUT       M00044	// ACK_PULSE 부저 ACK 상승 에지
; L39
LOAD      M00204	// HMI_COUNT_RESET CIMON 생산량 Reset: Manual Idle에서만 수락
AND NOT   M00054	// COUNT_RST_PREV 직전 스캔 HMI 생산량 Reset
AND NOT   F0009B
OUT       M00045	// COUNT_RST_PULSE 생산량 Reset 상승 에지
// 허가 조건 / 검사 응답
; L41
LOAD      M01000	// SIM_SAFE_OK 가상 안전 보조신호: 1=정상
AND       M01007	// SIM_DOOR_CLOSED 가상 문 닫힘 보조신호: 1=닫힘
OUT       M00001	// SAFE_MON_OK 안전 보조신호 정상: 가상 안전 및 문 닫힘
; L42
LOAD>=    D00100 20	// SEQ_STATE 현재 상태: 일반 조작에서 직접 쓰지 않음
AND<=     D00100 110	// SEQ_STATE 현재 상태: 일반 조작에서 직접 쓰지 않음
OUT       M00065	// CYCLE_ACTIVE 자동 사이클 중: 현재 상태 20~110
; L43
LOAD      M00065	// CYCLE_ACTIVE 자동 사이클 중: 현재 상태 20~110
AND<>     D00053 0	// MODE_SELECT 모드 선택: 0 Auto 1 Manual
OUT       M0004F	// MODE_ABORT 자동 사이클 중 Auto 이외 모드로 변경

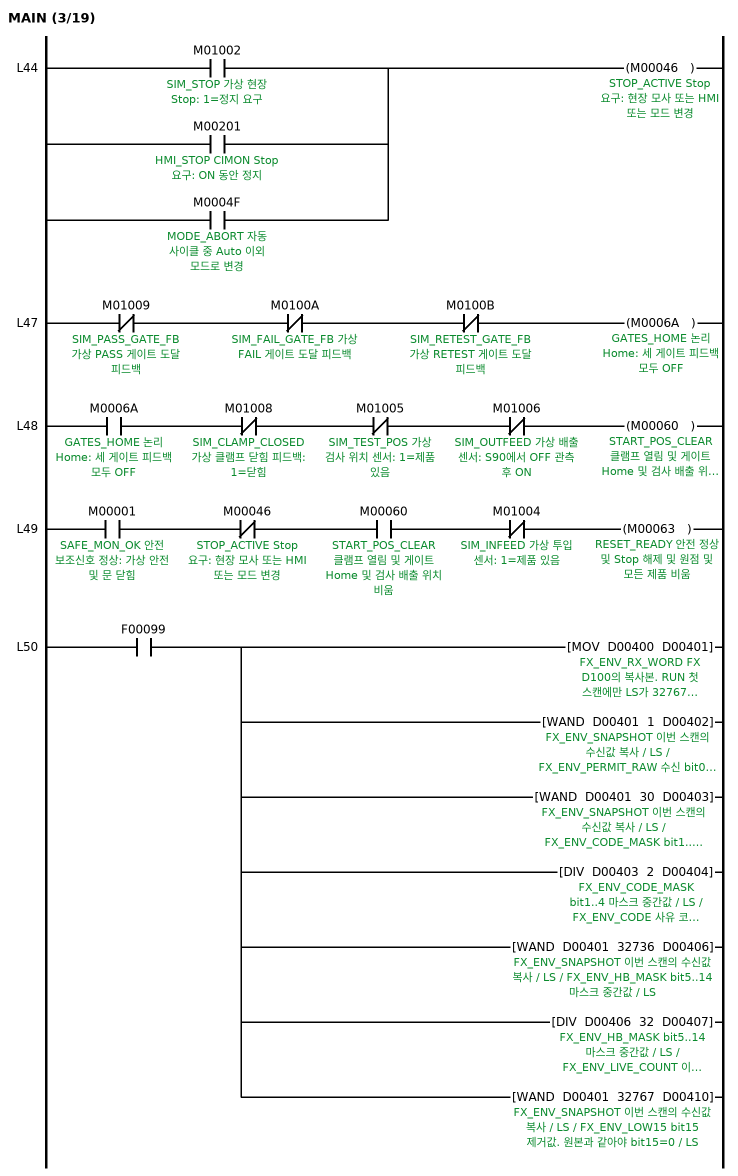
; L44
LOAD      M01002	// SIM_STOP 가상 현장 Stop: 1=정지 요구
OR        M00201	// HMI_STOP CIMON Stop 요구: ON 동안 정지
OR        M0004F	// MODE_ABORT 자동 사이클 중 Auto 이외 모드로 변경
OUT       M00046	// STOP_ACTIVE Stop 요구: 현장 모사 또는 HMI 또는 모드 변경
; L47
LOAD NOT  M01009	// SIM_PASS_GATE_FB 가상 PASS 게이트 도달 피드백
AND NOT   M0100A	// SIM_FAIL_GATE_FB 가상 FAIL 게이트 도달 피드백
AND NOT   M0100B	// SIM_RETEST_GATE_FB 가상 RETEST 게이트 도달 피드백
OUT       M0006A	// GATES_HOME 논리 Home: 세 게이트 피드백 모두 OFF
; L48
LOAD      M0006A	// GATES_HOME 논리 Home: 세 게이트 피드백 모두 OFF
AND NOT   M01008	// SIM_CLAMP_CLOSED 가상 클램프 닫힘 피드백: 1=닫힘
AND NOT   M01005	// SIM_TEST_POS 가상 검사 위치 센서: 1=제품 있음
AND NOT   M01006	// SIM_OUTFEED 가상 배출 센서: S90에서 OFF 관측 후 ON
OUT       M00060	// START_POS_CLEAR 클램프 열림 및 게이트 Home 및 검사 배출 위치 비움
; L49
LOAD      M00001	// SAFE_MON_OK 안전 보조신호 정상: 가상 안전 및 문 닫힘
AND NOT   M00046	// STOP_ACTIVE Stop 요구: 현장 모사 또는 HMI 또는 모드 변경
AND       M00060	// START_POS_CLEAR 클램프 열림 및 게이트 Home 및 검사 배출 위치 비움
AND NOT   M01004	// SIM_INFEED 가상 투입 센서: 1=제품 있음
OUT       M00063	// RESET_READY 안전 정상 및 Stop 해제 및 원점 및 모든 제품 비움
; L50
LOAD      F00099
MOV       D00400 D00401	// FX_ENV_RX_WORD FX D100의 복사본. RUN 첫 스캔에만 LS가 32767로 초기화. 이후 모의시험 작업자 또는 CIMON 한 곳이 기록 / FX_ENV_SNAPSHOT 이번 스캔의 수신값 복사 / LS
WAND      D00401 1 D00402	// FX_ENV_SNAPSHOT 이번 스캔의 수신값 복사 / LS / FX_ENV_PERMIT_RAW 수신 bit0, 0/1 / LS
WAND      D00401 30 D00403	// FX_ENV_SNAPSHOT 이번 스캔의 수신값 복사 / LS / FX_ENV_CODE_MASK bit1..4 마스크 중간값 / LS
DIV       D00403 2 D00404	// FX_ENV_CODE_MASK bit1..4 마스크 중간값 / LS / FX_ENV_CODE 사유 코드 0..15, 정상 형식은 0..6 / LS
WAND      D00401 32736 D00406	// FX_ENV_SNAPSHOT 이번 스캔의 수신값 복사 / LS / FX_ENV_HB_MASK bit5..14 마스크 중간값 / LS
DIV       D00406 32 D00407	// FX_ENV_HB_MASK bit5..14 마스크 중간값 / LS / FX_ENV_LIVE_COUNT 이번 카운터 0..1023 / LS
WAND      D00401 32767 D00410	// FX_ENV_SNAPSHOT 이번 스캔의 수신값 복사 / LS / FX_ENV_LOW15 bit15 제거값. 원본과 같아야 bit15=0 / LS

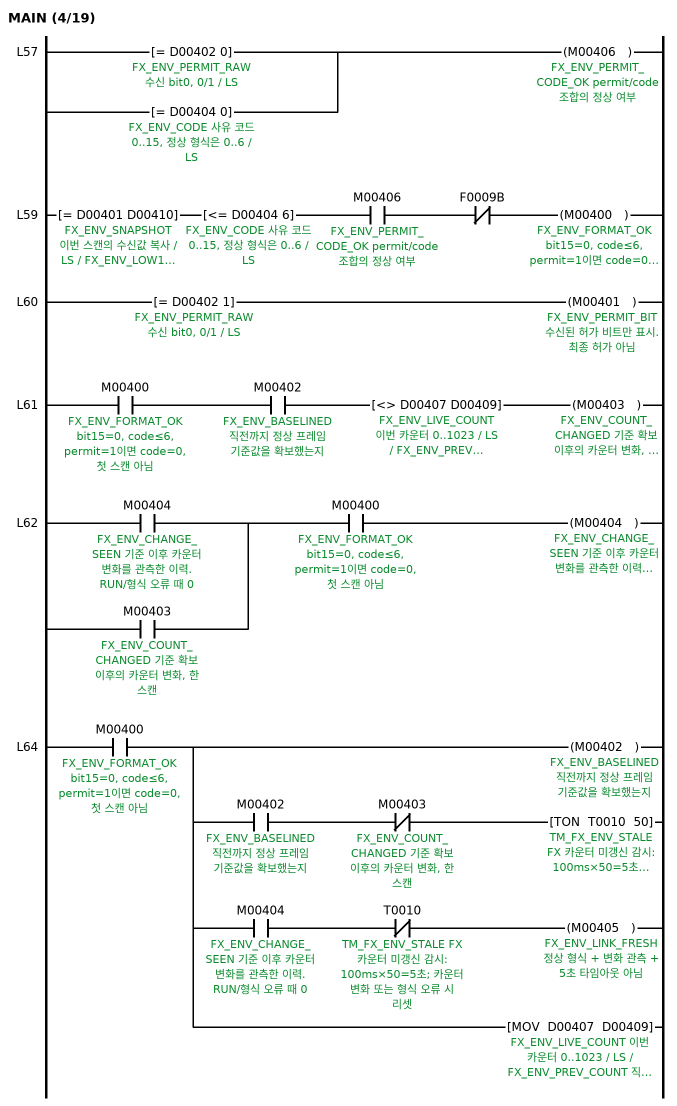
; L57
LOAD=     D00402 0	// FX_ENV_PERMIT_RAW 수신 bit0, 0/1 / LS
OR=       D00404 0	// FX_ENV_CODE 사유 코드 0..15, 정상 형식은 0..6 / LS
OUT       M00406	// FX_ENV_PERMIT_CODE_OK permit/code 조합의 정상 여부
; L59
LOAD=     D00401 D00410	// FX_ENV_SNAPSHOT 이번 스캔의 수신값 복사 / LS / FX_ENV_LOW15 bit15 제거값. 원본과 같아야 bit15=0 / LS
AND<=     D00404 6	// FX_ENV_CODE 사유 코드 0..15, 정상 형식은 0..6 / LS
AND       M00406	// FX_ENV_PERMIT_CODE_OK permit/code 조합의 정상 여부
AND NOT   F0009B
OUT       M00400	// FX_ENV_FORMAT_OK bit15=0, code≤6, permit=1이면 code=0, 첫 스캔 아님
; L60
LOAD=     D00402 1	// FX_ENV_PERMIT_RAW 수신 bit0, 0/1 / LS
OUT       M00401	// FX_ENV_PERMIT_BIT 수신된 허가 비트만 표시. 최종 허가 아님
; L61
LOAD      M00400	// FX_ENV_FORMAT_OK bit15=0, code≤6, permit=1이면 code=0, 첫 스캔 아님
AND       M00402	// FX_ENV_BASELINED 직전까지 정상 프레임 기준값을 확보했는지
AND<>     D00407 D00409	// FX_ENV_LIVE_COUNT 이번 카운터 0..1023 / LS / FX_ENV_PREV_COUNT 직전 정상 형식의 카운터 / LS
OUT       M00403	// FX_ENV_COUNT_CHANGED 기준 확보 이후의 카운터 변화, 한 스캔
; L62
LOAD      M00404	// FX_ENV_CHANGE_SEEN 기준 이후 카운터 변화를 관측한 이력. RUN/형식 오류 때 0
OR        M00403	// FX_ENV_COUNT_CHANGED 기준 확보 이후의 카운터 변화, 한 스캔
AND       M00400	// FX_ENV_FORMAT_OK bit15=0, code≤6, permit=1이면 code=0, 첫 스캔 아님
OUT       M00404	// FX_ENV_CHANGE_SEEN 기준 이후 카운터 변화를 관측한 이력. RUN/형식 오류 때 0
; L64
LOAD      M00400	// FX_ENV_FORMAT_OK bit15=0, code≤6, permit=1이면 code=0, 첫 스캔 아님
OUT       M00402	// FX_ENV_BASELINED 직전까지 정상 프레임 기준값을 확보했는지
MPUSH
AND       M00402	// FX_ENV_BASELINED 직전까지 정상 프레임 기준값을 확보했는지
AND NOT   M00403	// FX_ENV_COUNT_CHANGED 기준 확보 이후의 카운터 변화, 한 스캔
TON       T0010 50	// TM_FX_ENV_STALE FX 카운터 미갱신 감시: 100ms×50=5초; 카운터 변화 또는 형식 오류 시 리셋
MLOAD
AND       M00404	// FX_ENV_CHANGE_SEEN 기준 이후 카운터 변화를 관측한 이력. RUN/형식 오류 때 0
AND NOT   T0010	// TM_FX_ENV_STALE FX 카운터 미갱신 감시: 100ms×50=5초; 카운터 변화 또는 형식 오류 시 리셋
OUT       M00405	// FX_ENV_LINK_FRESH 정상 형식 + 변화 관측 + 5초 타임아웃 아님
MPOP
MOV       D00407 D00409	// FX_ENV_LIVE_COUNT 이번 카운터 0..1023 / LS / FX_ENV_PREV_COUNT 직전 정상 형식의 카운터 / LS

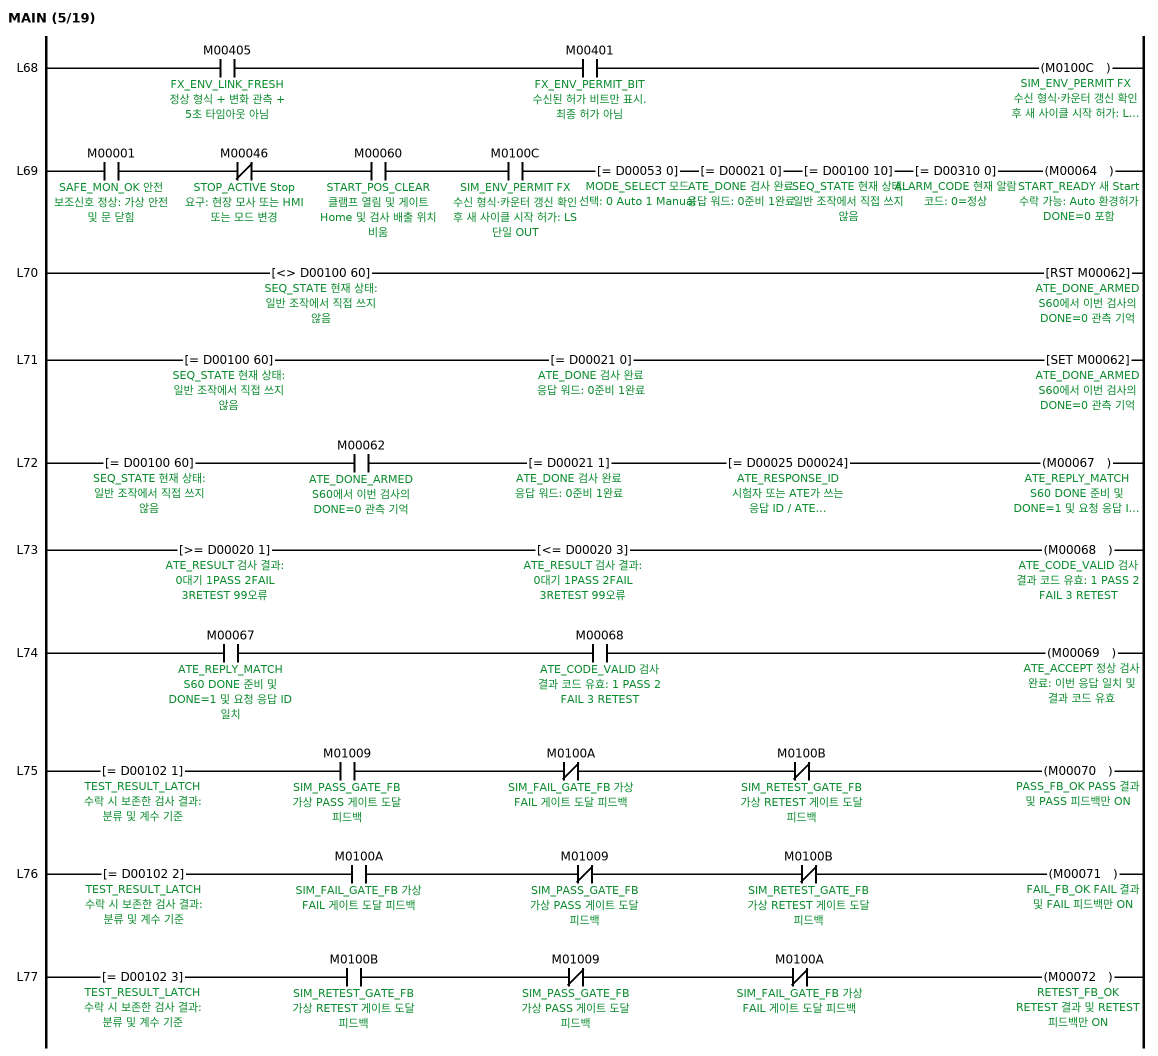
; L68
LOAD      M00405	// FX_ENV_LINK_FRESH 정상 형식 + 변화 관측 + 5초 타임아웃 아님
AND       M00401	// FX_ENV_PERMIT_BIT 수신된 허가 비트만 표시. 최종 허가 아님
OUT       M0100C	// SIM_ENV_PERMIT FX 수신 형식·카운터 갱신 확인 후 새 사이클 시작 허가: LS 단일 OUT
; L69
LOAD      M00001	// SAFE_MON_OK 안전 보조신호 정상: 가상 안전 및 문 닫힘
AND NOT   M00046	// STOP_ACTIVE Stop 요구: 현장 모사 또는 HMI 또는 모드 변경
AND       M00060	// START_POS_CLEAR 클램프 열림 및 게이트 Home 및 검사 배출 위치 비움
AND       M0100C	// SIM_ENV_PERMIT FX 수신 형식·카운터 갱신 확인 후 새 사이클 시작 허가: LS 단일 OUT
AND=      D00053 0	// MODE_SELECT 모드 선택: 0 Auto 1 Manual
AND=      D00021 0	// ATE_DONE 검사 완료 응답 워드: 0준비 1완료
AND=      D00100 10	// SEQ_STATE 현재 상태: 일반 조작에서 직접 쓰지 않음
AND=      D00310 0	// ALARM_CODE 현재 알람 코드: 0=정상
OUT       M00064	// START_READY 새 Start 수락 가능: Auto 환경허가 DONE=0 포함
; L70
LOAD<>    D00100 60	// SEQ_STATE 현재 상태: 일반 조작에서 직접 쓰지 않음
RST       M00062	// ATE_DONE_ARMED S60에서 이번 검사의 DONE=0 관측 기억
; L71
LOAD=     D00100 60	// SEQ_STATE 현재 상태: 일반 조작에서 직접 쓰지 않음
AND=      D00021 0	// ATE_DONE 검사 완료 응답 워드: 0준비 1완료
SET       M00062	// ATE_DONE_ARMED S60에서 이번 검사의 DONE=0 관측 기억
; L72
LOAD=     D00100 60	// SEQ_STATE 현재 상태: 일반 조작에서 직접 쓰지 않음
AND       M00062	// ATE_DONE_ARMED S60에서 이번 검사의 DONE=0 관측 기억
AND=      D00021 1	// ATE_DONE 검사 완료 응답 워드: 0준비 1완료
AND=      D00025 D00024	// ATE_RESPONSE_ID 시험자 또는 ATE가 쓰는 응답 ID / ATE_REQUEST_ID PLC 검사 요청 ID: 1~32000 RUN 초기화
OUT       M00067	// ATE_REPLY_MATCH S60 DONE 준비 및 DONE=1 및 요청 응답 ID 일치
; L73
LOAD>=    D00020 1	// ATE_RESULT 검사 결과: 0대기 1PASS 2FAIL 3RETEST 99오류
AND<=     D00020 3	// ATE_RESULT 검사 결과: 0대기 1PASS 2FAIL 3RETEST 99오류
OUT       M00068	// ATE_CODE_VALID 검사 결과 코드 유효: 1 PASS 2 FAIL 3 RETEST
; L74
LOAD      M00067	// ATE_REPLY_MATCH S60 DONE 준비 및 DONE=1 및 요청 응답 ID 일치
AND       M00068	// ATE_CODE_VALID 검사 결과 코드 유효: 1 PASS 2 FAIL 3 RETEST
OUT       M00069	// ATE_ACCEPT 정상 검사 완료: 이번 응답 일치 및 결과 코드 유효
; L75
LOAD=     D00102 1	// TEST_RESULT_LATCH 수락 시 보존한 검사 결과: 분류 및 계수 기준
AND       M01009	// SIM_PASS_GATE_FB 가상 PASS 게이트 도달 피드백
AND NOT   M0100A	// SIM_FAIL_GATE_FB 가상 FAIL 게이트 도달 피드백
AND NOT   M0100B	// SIM_RETEST_GATE_FB 가상 RETEST 게이트 도달 피드백
OUT       M00070	// PASS_FB_OK PASS 결과 및 PASS 피드백만 ON
; L76
LOAD=     D00102 2	// TEST_RESULT_LATCH 수락 시 보존한 검사 결과: 분류 및 계수 기준
AND       M0100A	// SIM_FAIL_GATE_FB 가상 FAIL 게이트 도달 피드백
AND NOT   M01009	// SIM_PASS_GATE_FB 가상 PASS 게이트 도달 피드백
AND NOT   M0100B	// SIM_RETEST_GATE_FB 가상 RETEST 게이트 도달 피드백
OUT       M00071	// FAIL_FB_OK FAIL 결과 및 FAIL 피드백만 ON
; L77
LOAD=     D00102 3	// TEST_RESULT_LATCH 수락 시 보존한 검사 결과: 분류 및 계수 기준
AND       M0100B	// SIM_RETEST_GATE_FB 가상 RETEST 게이트 도달 피드백
AND NOT   M01009	// SIM_PASS_GATE_FB 가상 PASS 게이트 도달 피드백
AND NOT   M0100A	// SIM_FAIL_GATE_FB 가상 FAIL 게이트 도달 피드백
OUT       M00072	// RETEST_FB_OK RETEST 결과 및 RETEST 피드백만 ON

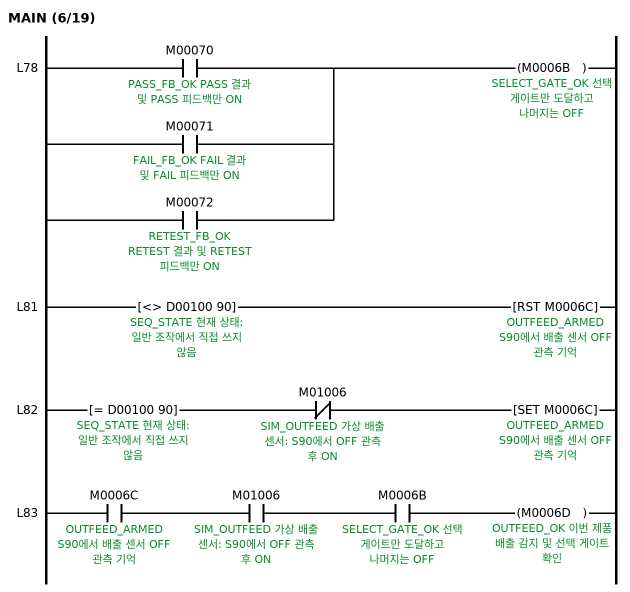
; L78
LOAD      M00070	// PASS_FB_OK PASS 결과 및 PASS 피드백만 ON
OR        M00071	// FAIL_FB_OK FAIL 결과 및 FAIL 피드백만 ON
OR        M00072	// RETEST_FB_OK RETEST 결과 및 RETEST 피드백만 ON
OUT       M0006B	// SELECT_GATE_OK 선택 게이트만 도달하고 나머지는 OFF
; L81
LOAD<>    D00100 90	// SEQ_STATE 현재 상태: 일반 조작에서 직접 쓰지 않음
RST       M0006C	// OUTFEED_ARMED S90에서 배출 센서 OFF 관측 기억
; L82
LOAD=     D00100 90	// SEQ_STATE 현재 상태: 일반 조작에서 직접 쓰지 않음
AND NOT   M01006	// SIM_OUTFEED 가상 배출 센서: S90에서 OFF 관측 후 ON
SET       M0006C	// OUTFEED_ARMED S90에서 배출 센서 OFF 관측 기억
; L83
LOAD      M0006C	// OUTFEED_ARMED S90에서 배출 센서 OFF 관측 기억
AND       M01006	// SIM_OUTFEED 가상 배출 센서: S90에서 OFF 관측 후 ON
AND       M0006B	// SELECT_GATE_OK 선택 게이트만 도달하고 나머지는 OFF
OUT       M0006D	// OUTFEED_OK 이번 제품 배출 감지 및 선택 게이트 확인

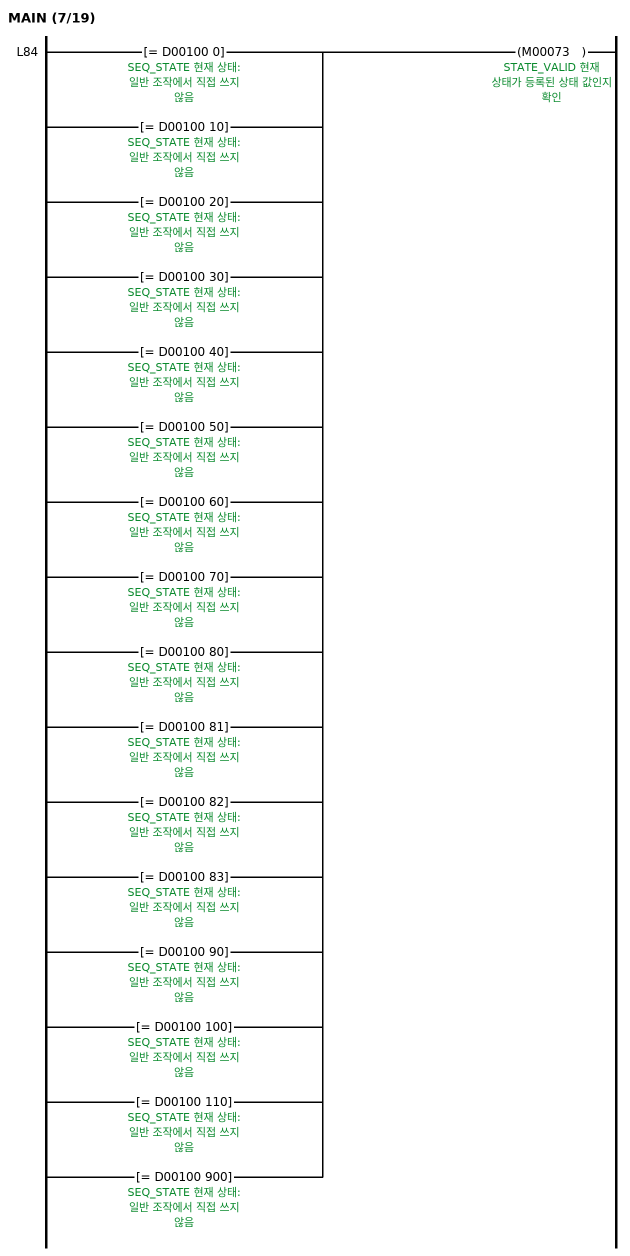
; L84
LOAD=     D00100 0	// SEQ_STATE 현재 상태: 일반 조작에서 직접 쓰지 않음
OR=       D00100 10	// SEQ_STATE 현재 상태: 일반 조작에서 직접 쓰지 않음
OR=       D00100 20	// SEQ_STATE 현재 상태: 일반 조작에서 직접 쓰지 않음
OR=       D00100 30	// SEQ_STATE 현재 상태: 일반 조작에서 직접 쓰지 않음
OR=       D00100 40	// SEQ_STATE 현재 상태: 일반 조작에서 직접 쓰지 않음
OR=       D00100 50	// SEQ_STATE 현재 상태: 일반 조작에서 직접 쓰지 않음
OR=       D00100 60	// SEQ_STATE 현재 상태: 일반 조작에서 직접 쓰지 않음
OR=       D00100 70	// SEQ_STATE 현재 상태: 일반 조작에서 직접 쓰지 않음
OR=       D00100 80	// SEQ_STATE 현재 상태: 일반 조작에서 직접 쓰지 않음
OR=       D00100 81	// SEQ_STATE 현재 상태: 일반 조작에서 직접 쓰지 않음
OR=       D00100 82	// SEQ_STATE 현재 상태: 일반 조작에서 직접 쓰지 않음
OR=       D00100 83	// SEQ_STATE 현재 상태: 일반 조작에서 직접 쓰지 않음
OR=       D00100 90	// SEQ_STATE 현재 상태: 일반 조작에서 직접 쓰지 않음
OR=       D00100 100	// SEQ_STATE 현재 상태: 일반 조작에서 직접 쓰지 않음
OR=       D00100 110	// SEQ_STATE 현재 상태: 일반 조작에서 직접 쓰지 않음
OR=       D00100 900	// SEQ_STATE 현재 상태: 일반 조작에서 직접 쓰지 않음
OUT       M00073	// STATE_VALID 현재 상태가 등록된 상태 값인지 확인

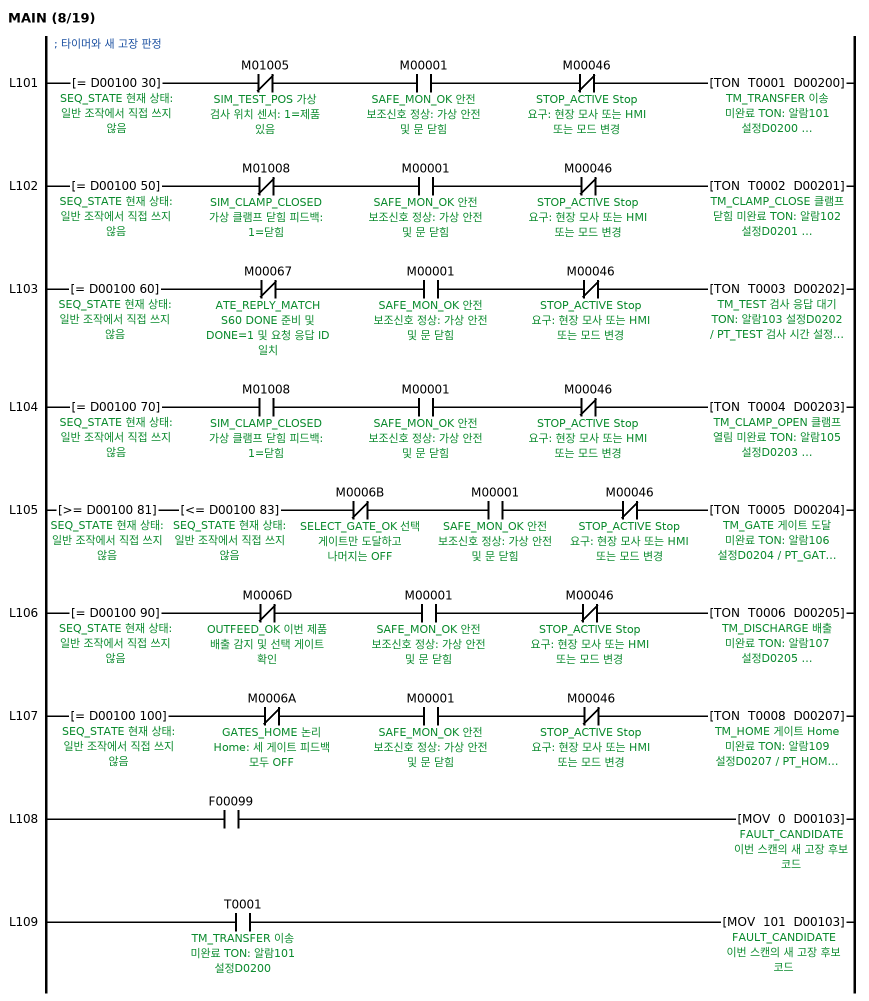
// 타이머와 새 고장 판정
; L101
LOAD=     D00100 30	// SEQ_STATE 현재 상태: 일반 조작에서 직접 쓰지 않음
AND NOT   M01005	// SIM_TEST_POS 가상 검사 위치 센서: 1=제품 있음
AND       M00001	// SAFE_MON_OK 안전 보조신호 정상: 가상 안전 및 문 닫힘
AND NOT   M00046	// STOP_ACTIVE Stop 요구: 현장 모사 또는 HMI 또는 모드 변경
TON       T0001 D00200	// TM_TRANSFER 이송 미완료 TON: 알람101 설정D0200 / PT_TRANSFER 이송 시간 설정: 100ms 단위 초기600=60초
; L102
LOAD=     D00100 50	// SEQ_STATE 현재 상태: 일반 조작에서 직접 쓰지 않음
AND NOT   M01008	// SIM_CLAMP_CLOSED 가상 클램프 닫힘 피드백: 1=닫힘
AND       M00001	// SAFE_MON_OK 안전 보조신호 정상: 가상 안전 및 문 닫힘
AND NOT   M00046	// STOP_ACTIVE Stop 요구: 현장 모사 또는 HMI 또는 모드 변경
TON       T0002 D00201	// TM_CLAMP_CLOSE 클램프 닫힘 미완료 TON: 알람102 설정D0201 / PT_CLAMP_CLOSE 클램프 닫힘 설정: 100ms 단위 초기600=60초
; L103
LOAD=     D00100 60	// SEQ_STATE 현재 상태: 일반 조작에서 직접 쓰지 않음
AND NOT   M00067	// ATE_REPLY_MATCH S60 DONE 준비 및 DONE=1 및 요청 응답 ID 일치
AND       M00001	// SAFE_MON_OK 안전 보조신호 정상: 가상 안전 및 문 닫힘
AND NOT   M00046	// STOP_ACTIVE Stop 요구: 현장 모사 또는 HMI 또는 모드 변경
TON       T0003 D00202	// TM_TEST 검사 응답 대기 TON: 알람103 설정D0202 / PT_TEST 검사 시간 설정: 100ms 단위 초기1200=120초
; L104
LOAD=     D00100 70	// SEQ_STATE 현재 상태: 일반 조작에서 직접 쓰지 않음
AND       M01008	// SIM_CLAMP_CLOSED 가상 클램프 닫힘 피드백: 1=닫힘
AND       M00001	// SAFE_MON_OK 안전 보조신호 정상: 가상 안전 및 문 닫힘
AND NOT   M00046	// STOP_ACTIVE Stop 요구: 현장 모사 또는 HMI 또는 모드 변경
TON       T0004 D00203	// TM_CLAMP_OPEN 클램프 열림 미완료 TON: 알람105 설정D0203 / PT_CLAMP_OPEN 클램프 열림 설정: 100ms 단위 초기600=60초
; L105
LOAD>=    D00100 81	// SEQ_STATE 현재 상태: 일반 조작에서 직접 쓰지 않음
AND<=     D00100 83	// SEQ_STATE 현재 상태: 일반 조작에서 직접 쓰지 않음
AND NOT   M0006B	// SELECT_GATE_OK 선택 게이트만 도달하고 나머지는 OFF
AND       M00001	// SAFE_MON_OK 안전 보조신호 정상: 가상 안전 및 문 닫힘
AND NOT   M00046	// STOP_ACTIVE Stop 요구: 현장 모사 또는 HMI 또는 모드 변경
TON       T0005 D00204	// TM_GATE 게이트 도달 미완료 TON: 알람106 설정D0204 / PT_GATE 게이트 도달 설정: 100ms 단위 초기600=60초
; L106
LOAD=     D00100 90	// SEQ_STATE 현재 상태: 일반 조작에서 직접 쓰지 않음
AND NOT   M0006D	// OUTFEED_OK 이번 제품 배출 감지 및 선택 게이트 확인
AND       M00001	// SAFE_MON_OK 안전 보조신호 정상: 가상 안전 및 문 닫힘
AND NOT   M00046	// STOP_ACTIVE Stop 요구: 현장 모사 또는 HMI 또는 모드 변경
TON       T0006 D00205	// TM_DISCHARGE 배출 미완료 TON: 알람107 설정D0205 / PT_DISCHARGE 배출 시간 설정: 100ms 단위 초기600=60초
; L107
LOAD=     D00100 100	// SEQ_STATE 현재 상태: 일반 조작에서 직접 쓰지 않음
AND NOT   M0006A	// GATES_HOME 논리 Home: 세 게이트 피드백 모두 OFF
AND       M00001	// SAFE_MON_OK 안전 보조신호 정상: 가상 안전 및 문 닫힘
AND NOT   M00046	// STOP_ACTIVE Stop 요구: 현장 모사 또는 HMI 또는 모드 변경
TON       T0008 D00207	// TM_HOME 게이트 Home 미완료 TON: 알람109 설정D0207 / PT_HOME Home 복귀 설정: 100ms 단위 초기600=60초
; L108
LOAD      F00099
MOV       0 D00103	// FAULT_CANDIDATE 이번 스캔의 새 고장 후보 코드
; L109
LOAD      T0001	// TM_TRANSFER 이송 미완료 TON: 알람101 설정D0200
MOV       101 D00103	// FAULT_CANDIDATE 이번 스캔의 새 고장 후보 코드

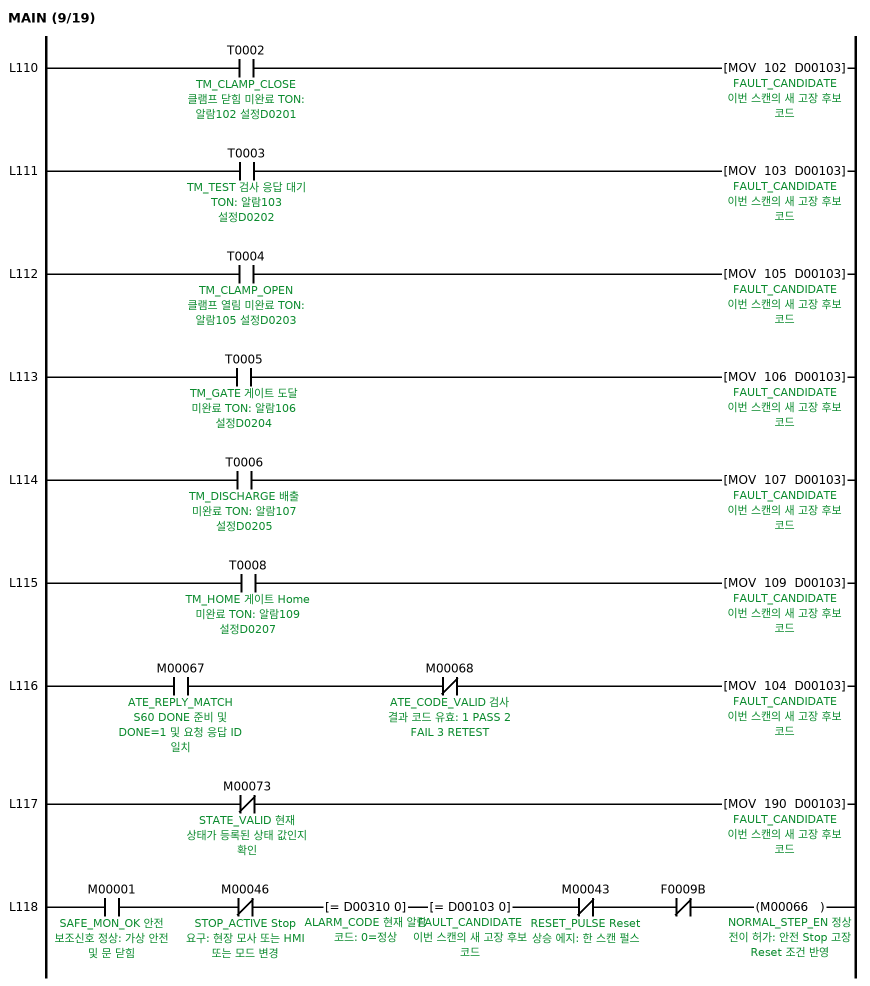
; L110
LOAD      T0002	// TM_CLAMP_CLOSE 클램프 닫힘 미완료 TON: 알람102 설정D0201
MOV       102 D00103	// FAULT_CANDIDATE 이번 스캔의 새 고장 후보 코드
; L111
LOAD      T0003	// TM_TEST 검사 응답 대기 TON: 알람103 설정D0202
MOV       103 D00103	// FAULT_CANDIDATE 이번 스캔의 새 고장 후보 코드
; L112
LOAD      T0004	// TM_CLAMP_OPEN 클램프 열림 미완료 TON: 알람105 설정D0203
MOV       105 D00103	// FAULT_CANDIDATE 이번 스캔의 새 고장 후보 코드
; L113
LOAD      T0005	// TM_GATE 게이트 도달 미완료 TON: 알람106 설정D0204
MOV       106 D00103	// FAULT_CANDIDATE 이번 스캔의 새 고장 후보 코드
; L114
LOAD      T0006	// TM_DISCHARGE 배출 미완료 TON: 알람107 설정D0205
MOV       107 D00103	// FAULT_CANDIDATE 이번 스캔의 새 고장 후보 코드
; L115
LOAD      T0008	// TM_HOME 게이트 Home 미완료 TON: 알람109 설정D0207
MOV       109 D00103	// FAULT_CANDIDATE 이번 스캔의 새 고장 후보 코드
; L116
LOAD      M00067	// ATE_REPLY_MATCH S60 DONE 준비 및 DONE=1 및 요청 응답 ID 일치
AND NOT   M00068	// ATE_CODE_VALID 검사 결과 코드 유효: 1 PASS 2 FAIL 3 RETEST
MOV       104 D00103	// FAULT_CANDIDATE 이번 스캔의 새 고장 후보 코드
; L117
LOAD NOT  M00073	// STATE_VALID 현재 상태가 등록된 상태 값인지 확인
MOV       190 D00103	// FAULT_CANDIDATE 이번 스캔의 새 고장 후보 코드
; L118
LOAD      M00001	// SAFE_MON_OK 안전 보조신호 정상: 가상 안전 및 문 닫힘
AND NOT   M00046	// STOP_ACTIVE Stop 요구: 현장 모사 또는 HMI 또는 모드 변경
AND=      D00310 0	// ALARM_CODE 현재 알람 코드: 0=정상
AND=      D00103 0	// FAULT_CANDIDATE 이번 스캔의 새 고장 후보 코드
AND NOT   M00043	// RESET_PULSE Reset 상승 에지: 한 스캔 펄스
AND NOT   F0009B
OUT       M00066	// NORMAL_STEP_EN 정상 전이 허가: 안전 Stop 고장 Reset 조건 반영

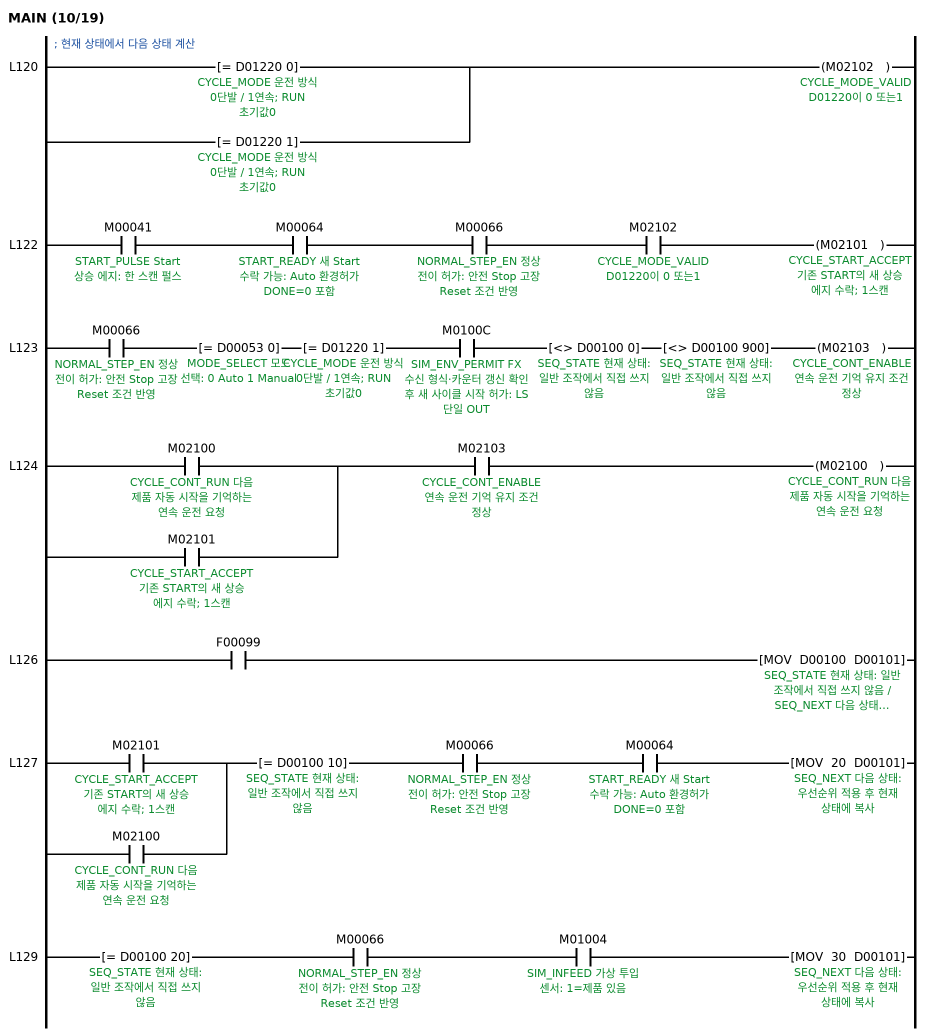
// 현재 상태에서 다음 상태 계산
; L120
LOAD=     D01220 0	// CYCLE_MODE 운전 방식 0단발 / 1연속; RUN 초기값0
OR=       D01220 1	// CYCLE_MODE 운전 방식 0단발 / 1연속; RUN 초기값0
OUT       M02102	// CYCLE_MODE_VALID D01220이 0 또는1
; L122
LOAD      M00041	// START_PULSE Start 상승 에지: 한 스캔 펄스
AND       M00064	// START_READY 새 Start 수락 가능: Auto 환경허가 DONE=0 포함
AND       M00066	// NORMAL_STEP_EN 정상 전이 허가: 안전 Stop 고장 Reset 조건 반영
AND       M02102	// CYCLE_MODE_VALID D01220이 0 또는1
OUT       M02101	// CYCLE_START_ACCEPT 기존 START의 새 상승 에지 수락; 1스캔
; L123
LOAD      M00066	// NORMAL_STEP_EN 정상 전이 허가: 안전 Stop 고장 Reset 조건 반영
AND=      D00053 0	// MODE_SELECT 모드 선택: 0 Auto 1 Manual
AND=      D01220 1	// CYCLE_MODE 운전 방식 0단발 / 1연속; RUN 초기값0
AND       M0100C	// SIM_ENV_PERMIT FX 수신 형식·카운터 갱신 확인 후 새 사이클 시작 허가: LS 단일 OUT
AND<>     D00100 0	// SEQ_STATE 현재 상태: 일반 조작에서 직접 쓰지 않음
AND<>     D00100 900	// SEQ_STATE 현재 상태: 일반 조작에서 직접 쓰지 않음
OUT       M02103	// CYCLE_CONT_ENABLE 연속 운전 기억 유지 조건 정상
; L124
LOAD      M02100	// CYCLE_CONT_RUN 다음 제품 자동 시작을 기억하는 연속 운전 요청
OR        M02101	// CYCLE_START_ACCEPT 기존 START의 새 상승 에지 수락; 1스캔
AND       M02103	// CYCLE_CONT_ENABLE 연속 운전 기억 유지 조건 정상
OUT       M02100	// CYCLE_CONT_RUN 다음 제품 자동 시작을 기억하는 연속 운전 요청
; L126
LOAD      F00099
MOV       D00100 D00101	// SEQ_STATE 현재 상태: 일반 조작에서 직접 쓰지 않음 / SEQ_NEXT 다음 상태: 우선순위 적용 후 현재 상태에 복사
; L127
LOAD      M02101	// CYCLE_START_ACCEPT 기존 START의 새 상승 에지 수락; 1스캔
OR        M02100	// CYCLE_CONT_RUN 다음 제품 자동 시작을 기억하는 연속 운전 요청
AND=      D00100 10	// SEQ_STATE 현재 상태: 일반 조작에서 직접 쓰지 않음
AND       M00066	// NORMAL_STEP_EN 정상 전이 허가: 안전 Stop 고장 Reset 조건 반영
AND       M00064	// START_READY 새 Start 수락 가능: Auto 환경허가 DONE=0 포함
MOV       20 D00101	// SEQ_NEXT 다음 상태: 우선순위 적용 후 현재 상태에 복사
; L129
LOAD=     D00100 20	// SEQ_STATE 현재 상태: 일반 조작에서 직접 쓰지 않음
AND       M00066	// NORMAL_STEP_EN 정상 전이 허가: 안전 Stop 고장 Reset 조건 반영
AND       M01004	// SIM_INFEED 가상 투입 센서: 1=제품 있음
MOV       30 D00101	// SEQ_NEXT 다음 상태: 우선순위 적용 후 현재 상태에 복사

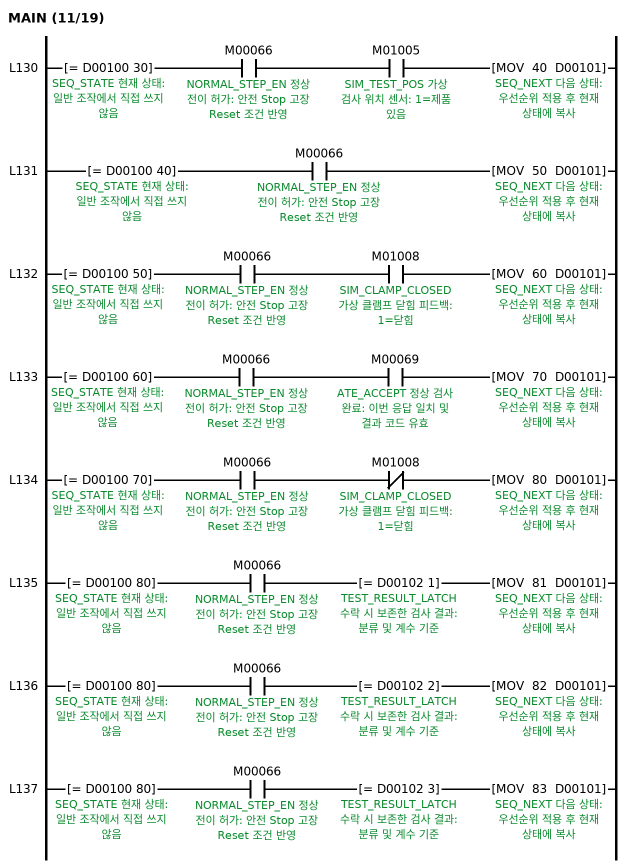
; L130
LOAD=     D00100 30	// SEQ_STATE 현재 상태: 일반 조작에서 직접 쓰지 않음
AND       M00066	// NORMAL_STEP_EN 정상 전이 허가: 안전 Stop 고장 Reset 조건 반영
AND       M01005	// SIM_TEST_POS 가상 검사 위치 센서: 1=제품 있음
MOV       40 D00101	// SEQ_NEXT 다음 상태: 우선순위 적용 후 현재 상태에 복사
; L131
LOAD=     D00100 40	// SEQ_STATE 현재 상태: 일반 조작에서 직접 쓰지 않음
AND       M00066	// NORMAL_STEP_EN 정상 전이 허가: 안전 Stop 고장 Reset 조건 반영
MOV       50 D00101	// SEQ_NEXT 다음 상태: 우선순위 적용 후 현재 상태에 복사
; L132
LOAD=     D00100 50	// SEQ_STATE 현재 상태: 일반 조작에서 직접 쓰지 않음
AND       M00066	// NORMAL_STEP_EN 정상 전이 허가: 안전 Stop 고장 Reset 조건 반영
AND       M01008	// SIM_CLAMP_CLOSED 가상 클램프 닫힘 피드백: 1=닫힘
MOV       60 D00101	// SEQ_NEXT 다음 상태: 우선순위 적용 후 현재 상태에 복사
; L133
LOAD=     D00100 60	// SEQ_STATE 현재 상태: 일반 조작에서 직접 쓰지 않음
AND       M00066	// NORMAL_STEP_EN 정상 전이 허가: 안전 Stop 고장 Reset 조건 반영
AND       M00069	// ATE_ACCEPT 정상 검사 완료: 이번 응답 일치 및 결과 코드 유효
MOV       70 D00101	// SEQ_NEXT 다음 상태: 우선순위 적용 후 현재 상태에 복사
; L134
LOAD=     D00100 70	// SEQ_STATE 현재 상태: 일반 조작에서 직접 쓰지 않음
AND       M00066	// NORMAL_STEP_EN 정상 전이 허가: 안전 Stop 고장 Reset 조건 반영
AND NOT   M01008	// SIM_CLAMP_CLOSED 가상 클램프 닫힘 피드백: 1=닫힘
MOV       80 D00101	// SEQ_NEXT 다음 상태: 우선순위 적용 후 현재 상태에 복사
; L135
LOAD=     D00100 80	// SEQ_STATE 현재 상태: 일반 조작에서 직접 쓰지 않음
AND       M00066	// NORMAL_STEP_EN 정상 전이 허가: 안전 Stop 고장 Reset 조건 반영
AND=      D00102 1	// TEST_RESULT_LATCH 수락 시 보존한 검사 결과: 분류 및 계수 기준
MOV       81 D00101	// SEQ_NEXT 다음 상태: 우선순위 적용 후 현재 상태에 복사
; L136
LOAD=     D00100 80	// SEQ_STATE 현재 상태: 일반 조작에서 직접 쓰지 않음
AND       M00066	// NORMAL_STEP_EN 정상 전이 허가: 안전 Stop 고장 Reset 조건 반영
AND=      D00102 2	// TEST_RESULT_LATCH 수락 시 보존한 검사 결과: 분류 및 계수 기준
MOV       82 D00101	// SEQ_NEXT 다음 상태: 우선순위 적용 후 현재 상태에 복사
; L137
LOAD=     D00100 80	// SEQ_STATE 현재 상태: 일반 조작에서 직접 쓰지 않음
AND       M00066	// NORMAL_STEP_EN 정상 전이 허가: 안전 Stop 고장 Reset 조건 반영
AND=      D00102 3	// TEST_RESULT_LATCH 수락 시 보존한 검사 결과: 분류 및 계수 기준
MOV       83 D00101	// SEQ_NEXT 다음 상태: 우선순위 적용 후 현재 상태에 복사

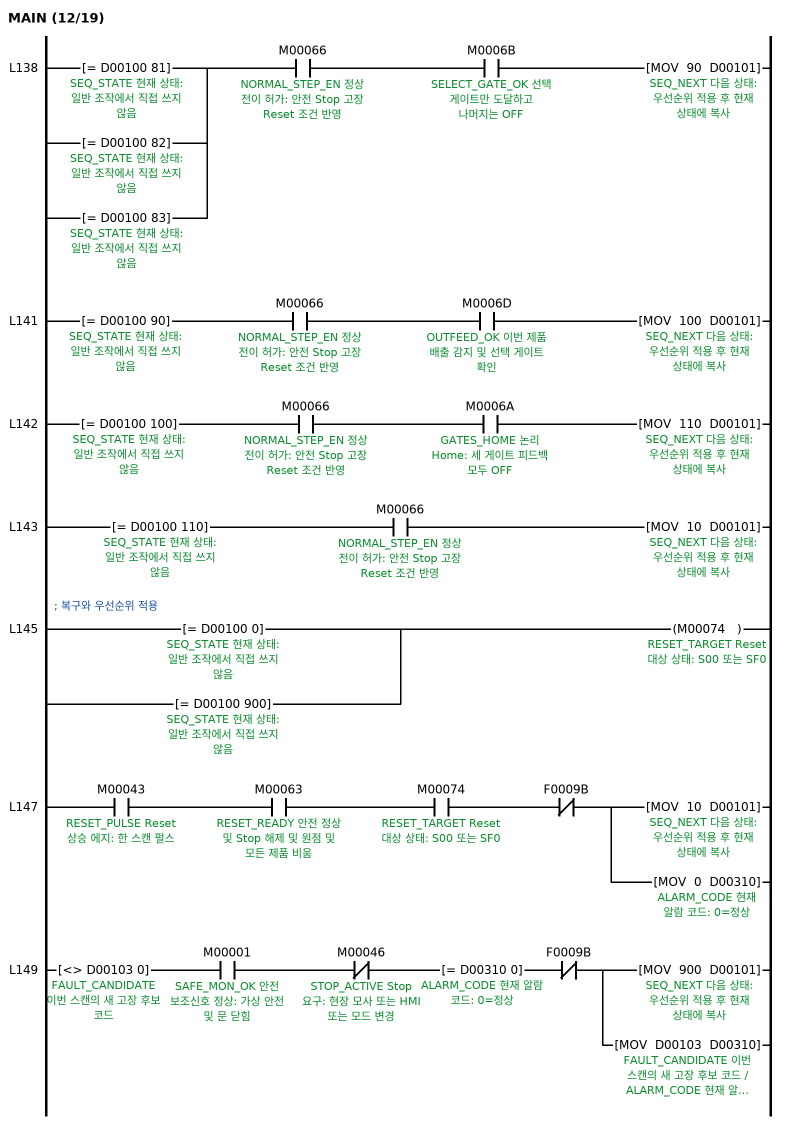
; L138
LOAD=     D00100 81	// SEQ_STATE 현재 상태: 일반 조작에서 직접 쓰지 않음
OR=       D00100 82	// SEQ_STATE 현재 상태: 일반 조작에서 직접 쓰지 않음
OR=       D00100 83	// SEQ_STATE 현재 상태: 일반 조작에서 직접 쓰지 않음
AND       M00066	// NORMAL_STEP_EN 정상 전이 허가: 안전 Stop 고장 Reset 조건 반영
AND       M0006B	// SELECT_GATE_OK 선택 게이트만 도달하고 나머지는 OFF
MOV       90 D00101	// SEQ_NEXT 다음 상태: 우선순위 적용 후 현재 상태에 복사
; L141
LOAD=     D00100 90	// SEQ_STATE 현재 상태: 일반 조작에서 직접 쓰지 않음
AND       M00066	// NORMAL_STEP_EN 정상 전이 허가: 안전 Stop 고장 Reset 조건 반영
AND       M0006D	// OUTFEED_OK 이번 제품 배출 감지 및 선택 게이트 확인
MOV       100 D00101	// SEQ_NEXT 다음 상태: 우선순위 적용 후 현재 상태에 복사
; L142
LOAD=     D00100 100	// SEQ_STATE 현재 상태: 일반 조작에서 직접 쓰지 않음
AND       M00066	// NORMAL_STEP_EN 정상 전이 허가: 안전 Stop 고장 Reset 조건 반영
AND       M0006A	// GATES_HOME 논리 Home: 세 게이트 피드백 모두 OFF
MOV       110 D00101	// SEQ_NEXT 다음 상태: 우선순위 적용 후 현재 상태에 복사
; L143
LOAD=     D00100 110	// SEQ_STATE 현재 상태: 일반 조작에서 직접 쓰지 않음
AND       M00066	// NORMAL_STEP_EN 정상 전이 허가: 안전 Stop 고장 Reset 조건 반영
MOV       10 D00101	// SEQ_NEXT 다음 상태: 우선순위 적용 후 현재 상태에 복사
// 복구와 우선순위 적용
; L145
LOAD=     D00100 0	// SEQ_STATE 현재 상태: 일반 조작에서 직접 쓰지 않음
OR=       D00100 900	// SEQ_STATE 현재 상태: 일반 조작에서 직접 쓰지 않음
OUT       M00074	// RESET_TARGET Reset 대상 상태: S00 또는 SF0
; L147
LOAD      M00043	// RESET_PULSE Reset 상승 에지: 한 스캔 펄스
AND       M00063	// RESET_READY 안전 정상 및 Stop 해제 및 원점 및 모든 제품 비움
AND       M00074	// RESET_TARGET Reset 대상 상태: S00 또는 SF0
AND NOT   F0009B
MOV       10 D00101	// SEQ_NEXT 다음 상태: 우선순위 적용 후 현재 상태에 복사
MOV       0 D00310	// ALARM_CODE 현재 알람 코드: 0=정상
; L149
LOAD<>    D00103 0	// FAULT_CANDIDATE 이번 스캔의 새 고장 후보 코드
AND       M00001	// SAFE_MON_OK 안전 보조신호 정상: 가상 안전 및 문 닫힘
AND NOT   M00046	// STOP_ACTIVE Stop 요구: 현장 모사 또는 HMI 또는 모드 변경
AND=      D00310 0	// ALARM_CODE 현재 알람 코드: 0=정상
AND NOT   F0009B
MOV       900 D00101	// SEQ_NEXT 다음 상태: 우선순위 적용 후 현재 상태에 복사
MOV       D00103 D00310	// FAULT_CANDIDATE 이번 스캔의 새 고장 후보 코드 / ALARM_CODE 현재 알람 코드: 0=정상

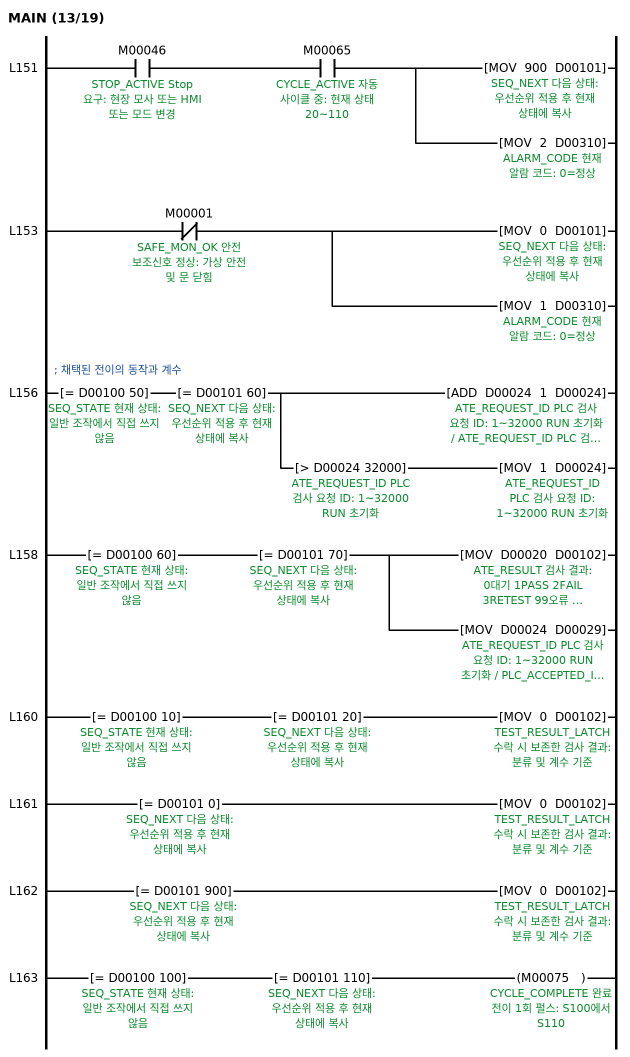
; L151
LOAD      M00046	// STOP_ACTIVE Stop 요구: 현장 모사 또는 HMI 또는 모드 변경
AND       M00065	// CYCLE_ACTIVE 자동 사이클 중: 현재 상태 20~110
MOV       900 D00101	// SEQ_NEXT 다음 상태: 우선순위 적용 후 현재 상태에 복사
MOV       2 D00310	// ALARM_CODE 현재 알람 코드: 0=정상
; L153
LOAD NOT  M00001	// SAFE_MON_OK 안전 보조신호 정상: 가상 안전 및 문 닫힘
MOV       0 D00101	// SEQ_NEXT 다음 상태: 우선순위 적용 후 현재 상태에 복사
MOV       1 D00310	// ALARM_CODE 현재 알람 코드: 0=정상
// 채택된 전이의 동작과 계수
; L156
LOAD=     D00100 50	// SEQ_STATE 현재 상태: 일반 조작에서 직접 쓰지 않음
AND=      D00101 60	// SEQ_NEXT 다음 상태: 우선순위 적용 후 현재 상태에 복사
ADD       D00024 1 D00024	// ATE_REQUEST_ID PLC 검사 요청 ID: 1~32000 RUN 초기화 / ATE_REQUEST_ID PLC 검사 요청 ID: 1~32000 RUN 초기화
AND>      D00024 32000	// ATE_REQUEST_ID PLC 검사 요청 ID: 1~32000 RUN 초기화
MOV       1 D00024	// ATE_REQUEST_ID PLC 검사 요청 ID: 1~32000 RUN 초기화
; L158
LOAD=     D00100 60	// SEQ_STATE 현재 상태: 일반 조작에서 직접 쓰지 않음
AND=      D00101 70	// SEQ_NEXT 다음 상태: 우선순위 적용 후 현재 상태에 복사
MOV       D00020 D00102	// ATE_RESULT 검사 결과: 0대기 1PASS 2FAIL 3RETEST 99오류 / TEST_RESULT_LATCH 수락 시 보존한 검사 결과: 분류 및 계수 기준
MOV       D00024 D00029	// ATE_REQUEST_ID PLC 검사 요청 ID: 1~32000 RUN 초기화 / PLC_ACCEPTED_ID 상태 60→70이 최종 채택될 때 D00024를 보존한 번호
; L160
LOAD=     D00100 10	// SEQ_STATE 현재 상태: 일반 조작에서 직접 쓰지 않음
AND=      D00101 20	// SEQ_NEXT 다음 상태: 우선순위 적용 후 현재 상태에 복사
MOV       0 D00102	// TEST_RESULT_LATCH 수락 시 보존한 검사 결과: 분류 및 계수 기준
; L161
LOAD=     D00101 0	// SEQ_NEXT 다음 상태: 우선순위 적용 후 현재 상태에 복사
MOV       0 D00102	// TEST_RESULT_LATCH 수락 시 보존한 검사 결과: 분류 및 계수 기준
; L162
LOAD=     D00101 900	// SEQ_NEXT 다음 상태: 우선순위 적용 후 현재 상태에 복사
MOV       0 D00102	// TEST_RESULT_LATCH 수락 시 보존한 검사 결과: 분류 및 계수 기준
; L163
LOAD=     D00100 100	// SEQ_STATE 현재 상태: 일반 조작에서 직접 쓰지 않음
AND=      D00101 110	// SEQ_NEXT 다음 상태: 우선순위 적용 후 현재 상태에 복사
OUT       M00075	// CYCLE_COMPLETE 완료 전이 1회 펄스: S100에서 S110

